{region 'Documentation'}
(*!
<summary>No asynchronous test resource remains to stop.</summary>
*)
{endregion}
METHOD PROTECTED ProcessAbort
VAR_INPUT
    Enable : BOOL; //! Phase permission supplied by the owning Test Case; FALSE does not authorize progression, while observation may continue.
END_VAR
IF Enable THEN
    CompleteAbort();
END_IF;
END_METHOD

{region 'Documentation'}
(*!
<summary>Evaluates each scripted call before the test advances; failures remain latched across both runs.</summary>
*)
{endregion}
METHOD PROTECTED ProcessAssertions
VAR_INPUT
    Enable : BOOL; //! Phase permission supplied by the owning Test Case; FALSE does not authorize progression, while observation may continue.
END_VAR
FStatePath(Enable := Enable,
    State := State,
    IN := FStatePathMatches);
FTaskMapping(Enable := Enable,
    State := State,
    IN := FTaskMappingMatches);
FOwnerResult(Enable := Enable,
    State := State,
    IN := FOwnerResultMatches);
FStatusCounters(Enable := Enable,
    State := State,
    IN := FStatusCountersMatches);
FCallOrder(Enable := Enable,
    State := State,
    IN := FCallOrderMatches);
FReadiness(Enable := Enable,
    State := State,
    IN := FReadinessMatches);
FFinalEvents(Enable := Enable,
    State := State,
    IN := FFinalEventsMatches);
FAggregationPayload(Enable := Enable,
    State := State,
    IN := FAggregationPayloadMatches);
FCaptureIntegrity(Enable := Enable,
    State := State,
    IN := FCaptureIntegrityMatches);
IF Enable THEN
    FStepChecked := TRUE;
END_IF;
END_METHOD

{region 'Documentation'}
(*!
<summary>No resource Preparation is required for this controlled owner scenario.</summary>
*)
{endregion}
METHOD PROTECTED ProcessPreparations
VAR_INPUT
    // SA0033: Required override; the scenario has no Preparation phase.
    {attribute 'analysis' := '-33'}
    Enable : BOOL; //! Phase permission supplied by the owning Test Case; FALSE does not authorize progression, while observation may continue.
END_VAR
END_METHOD

{region 'Documentation'}
(*!
<summary>Restarts the test script and clears checking Assertions; subject setup belongs to the next test attempt.</summary>
*)
{endregion}
METHOD PROTECTED ProcessReset
FStep := Setup;
FRun := 1;
FStepChecked := FALSE;
FStatePathMatches := TRUE;
FTaskMappingMatches := TRUE;
FOwnerResultMatches := TRUE;
FStatusCountersMatches := TRUE;
FCallOrderMatches := TRUE;
FReadinessMatches := TRUE;
FFinalEventsMatches := TRUE;
FAggregationPayloadMatches := TRUE;
FCaptureIntegrityMatches := TRUE;
FStatePath.Reset();
FTaskMapping.Reset();
FOwnerResult.Reset();
FStatusCounters.Reset();
FCallOrder.Reset();
FReadiness.Reset();
FFinalEvents.Reset();
FAggregationPayload.Reset();
FCaptureIntegrity.Reset();
CompleteReset();
END_METHOD

{region 'Documentation'}
(*!
<summary>Advances the explicit test script with at most one subject FB call per active PLC cycle.</summary>
*)
{endregion}
METHOD PROTECTED ProcessTests
VAR_INPUT
    Enable : BOOL; //! Phase permission supplied by the owning Test Case; FALSE does not authorize progression, while observation may continue.
END_VAR
IF NOT Enable THEN
    RETURN;
END_IF;
IF FStepChecked THEN
    IF FStep = StartWithoutReset THEN
        IF FRun = RunCount THEN
            CompleteTests();
            RETURN;
        END_IF;
        FRun := FRun + 1;
        FStep := Setup;
    ELSE
        FStep := FStep + 1;
    END_IF;
    FStepChecked := FALSE;
    NextTestState();
END_IF;
RunStep();
END_METHOD

{region 'Documentation'}
(*!
<summary>Arranges one root cycle, executes it once and compares state, counters and call ordering.</summary>
*)
{endregion}
METHOD PRIVATE RunStep
VAR
    Config : ST_RunConfig;
    FirstView : ST_OrchestrationObservation;
    SecondView : ST_OrchestrationObservation;
    ExpectedState : E_State;
    ExpectedTask : E_OrchestratorTask;
    ExpectedResult : E_Result := E_Result.NotEvaluated;
    ExpectedReady : BOOL;
    ExpectedIdleCount : UINT;
    ExpectedRunningCount : UINT;
    ExpectedCompletedCount : UINT;
    ExpectedPassedCount : UINT;
    ExpectedFailedCount : UINT;
    ExpectedExecutionStatus : E_ExecutionStatus;
    FirstChild : I_Orchestratable;
    LastChild : I_Orchestratable;
    FirstStateBeforeCall : E_State;
    LastStateBeforeCall : E_State;
    Snapshot : ST_RunControlStatus;
    ExpectedCalls : UINT;
END_VAR
CASE FStep OF
    Setup:
        FRunChildResult := E_Result.Passed;
        IF FRun = 1 THEN
            FRunChildResult := FirstChildResult;
            IF NOT FCapture.Initialize(Buffer := FEvents,
                FifoControl := FCaptureFifo,
                Status := FCaptureStatus) THEN
                Error(Message := 'Root lifecycle capture could not be initialized.');
                RETURN;
            END_IF;
            Config.CompletionDelay := T#0ms;
            FHelper.BeginScenario();
            FSubject.Bind(Publisher := FCapture,
                Helper := FHelper,
                Config := Config);
            IF NOT FSubject.Initialize(Name := 'LifecycleSubject',
                EventBuffer := FCapture) THEN
                Error(Message := 'Root lifecycle subject could not be initialized.');
                RETURN;
            END_IF;
        ELSE
            FHelper.SetObservation(Ready := FALSE);
            FSubject.RequestReset();
        END_IF;
        FirstView.State := E_State.Reset;
        FirstView.Ready := FALSE;
        SecondView := FirstView;
        ExpectedState := E_State.Reset;
        ExpectedTask := E_OrchestratorTask.Reset;
        ExpectedExecutionStatus := E_ExecutionStatus.Reset;

    ChildrenReady:
        ExpectedState := E_State.Reset;
        ExpectedTask := E_OrchestratorTask.Reset;
        ExpectedExecutionStatus := E_ExecutionStatus.Reset;
        ExpectedIdleCount := ExpectedChildCount;

    ResetFinished:
        FHelper.SetObservation(Ready := FALSE,
            ResetFinished := TRUE);
        ExpectedState := E_State.Idle;
        ExpectedTask := E_OrchestratorTask.Idle;
        ExpectedExecutionStatus := E_ExecutionStatus.Idle;
        ExpectedIdleCount := ExpectedChildCount;

    StartReady:
        FHelper.SetObservation(Ready := TRUE);
        ExpectedState := E_State.Idle;
        ExpectedTask := E_OrchestratorTask.Idle;
        ExpectedExecutionStatus := E_ExecutionStatus.Idle;
        ExpectedIdleCount := ExpectedChildCount;
        ExpectedReady := TRUE;

    StartRequested:
        FSubject.RequestStart();
        FirstView.State := E_State.Running;
        FirstView.Ready := FALSE;
        ExpectedState := E_State.Starting;
        ExpectedTask := E_OrchestratorTask.Execution;
        ExpectedExecutionStatus := E_ExecutionStatus.Starting;
        ExpectedIdleCount := 1;
        ExpectedRunningCount := 1;

    FirstChildCompleted:
        FHelper.SetObservation(Ready := FALSE);
        FirstView.State := E_State.Completed;
        FirstView.Result := FRunChildResult;
        FirstView.Ready := FALSE;
        FirstView.Complete := TRUE;
        SecondView.State := E_State.Running;
        SecondView.Ready := FALSE;
        ExpectedState := E_State.Running;
        ExpectedTask := E_OrchestratorTask.Execution;
        ExpectedExecutionStatus := E_ExecutionStatus.Running;
        ExpectedRunningCount := 1;
        ExpectedCompletedCount := 1;
        ExpectedFailedCount := BOOL_TO_UINT(FRunChildResult = E_Result.Failed);
        ExpectedPassedCount := 1 - ExpectedFailedCount;

    AllChildrenCompleted, WaitForHelper, OwnerCompleting, OwnerCompleted, HoldCompleted, StartWithoutReset:
        FHelper.SetObservation(Ready := FALSE);
        FirstView.State := E_State.Completed;
        FirstView.Result := FRunChildResult;
        FirstView.Ready := FALSE;
        FirstView.Complete := TRUE;
        SecondView := FirstView;
        SecondView.Result := E_Result.Passed;
        ExpectedTask := E_OrchestratorTask.Execution;
        ExpectedCompletedCount := ExpectedChildCount;
        ExpectedFailedCount := BOOL_TO_UINT(FRunChildResult = E_Result.Failed);
        ExpectedPassedCount := ExpectedChildCount - ExpectedFailedCount;
        CASE FStep OF
            AllChildrenCompleted, WaitForHelper:
                ExpectedState := E_State.Running;
                ExpectedExecutionStatus := E_ExecutionStatus.Running;
            OwnerCompleting:
                FHelper.SetObservation(Ready := FALSE,
                    ExecutionFinished := TRUE);
                ExpectedState := E_State.Completing;
                ExpectedExecutionStatus := E_ExecutionStatus.Completing;
                ExpectedResult := FRunChildResult;
        ELSE
            IF FStep = StartWithoutReset THEN
                FSubject.RequestStart();
            END_IF;
            ExpectedState := E_State.Completed;
            ExpectedTask := E_OrchestratorTask.Idle;
            ExpectedExecutionStatus := E_ExecutionStatus.Completed;
            ExpectedResult := FRunChildResult;
        END_CASE;
ELSE
    Error(Message := 'Unexpected root lifecycle test step.');
    RETURN;
END_CASE;

FirstChild := FSubject.GetChild(Index := FSubject.ChildArrayLowerBound);
LastChild := FSubject.GetChild(Index := FSubject.ChildArrayLowerBound + UINT_TO_DINT(FSubject.ChildCount) - 1);
FirstStateBeforeCall := FirstChild.State;
LastStateBeforeCall := LastChild.State;
FSubject.SetChildObservations(FirstChild := FirstView,
    SecondChild := SecondView);
FSubject(ControlData := FControl);
Snapshot := FSubject.Status;
ExpectedCalls := INT_TO_UINT((FRun - 1) * StepsPerRun + FStep + 1);

FStatePathMatches := (FSubject.State = ExpectedState)
    AND (Snapshot.Execution.State = ExpectedState)
    AND (Snapshot.Execution.ExecutionStatus = ExpectedExecutionStatus)
    AND (FControl.Status.Execution.State = ExpectedState)
    AND (FControl.Name = 'LifecycleSubject');
FTaskMappingMatches := FHelper.CurrentTask = ExpectedTask;
FOwnerResultMatches := (FSubject.Result = ExpectedResult)
    AND (Snapshot.Execution.Result = ExpectedResult)
    AND (FControl.Status.Execution.Result = ExpectedResult)
    AND NOT FSubject.HasError;
FStatusCountersMatches := (Snapshot.SuiteCountTotal = ExpectedChildCount)
    AND (Snapshot.SuiteCountIdle = ExpectedIdleCount)
    AND (Snapshot.SuiteCountRunning = ExpectedRunningCount)
    AND (Snapshot.SuiteCountCompleted = ExpectedCompletedCount)
    AND (Snapshot.SuiteCountPassed = ExpectedPassedCount)
    AND (Snapshot.SuiteCountFailed = ExpectedFailedCount)
    AND (Snapshot.SuiteCountError = 0) AND (Snapshot.SuiteCountInactive = 0)
    AND (FControl.Status.SuiteCountIdle = ExpectedIdleCount)
    AND (FControl.Status.SuiteCountRunning = ExpectedRunningCount)
    AND (FControl.Status.SuiteCountCompleted = ExpectedCompletedCount)
    AND (FControl.Status.SuiteCountPassed = ExpectedPassedCount)
    AND (FControl.Status.SuiteCountFailed = ExpectedFailedCount);
FCallOrderMatches := (FHelper.InitializeCount = 1) AND (FSubject.ConfigureCount = 1)
    AND (FHelper.ExecuteCount = ExpectedCalls)
    AND (FSubject.ChildCallCount = ExpectedCalls)
    AND FSubject.ChildBodyCallsMatch
    AND (FHelper.FirstChildStateAtExecute = FirstStateBeforeCall)
    AND (FHelper.LastChildStateAtExecute = LastStateBeforeCall)
    AND (FirstChild.State = FirstView.State) AND (LastChild.State = SecondView.State);
FReadinessMatches := (FSubject.IsReady = ExpectedReady)
    AND (Snapshot.Execution.Ready = ExpectedReady)
    AND (FSubject.IsComplete = (ExpectedState = E_State.Completed));
FCaptureIntegrityMatches := (FCaptureStatus.LostEventCount = 0)
    AND (FCaptureFifo.ElementCount = FCaptureStatus.SequenceId);
IF FStep = Setup THEN
    FOwnerResultMatches := FOwnerResultMatches AND (Snapshot.Runtime = T#0ms);
END_IF;
IF FStep = OwnerCompleting THEN
    FRunRuntime[FRun] := Snapshot.Runtime;
END_IF;
CheckFinalEvents();
END_METHOD

END_FUNCTION_BLOCK

// ---- SelfTests/TestCases/TestSuite_RunControlLifecycle/Test_RunControlRequests.TcPOU
{region 'Documentation'}
(*!
<summary>Checks direct root requests, one-call consumption and Reset/Abort/Start priority.</summary>
<description>
The controlled helper only supplies readiness and completion. The script covers a Start
received while not ready, repeated Start method calls before one FB call, Start while active,
Abort together with Start, and Reset together with both lower-priority requests.
A repeated Reset while already resetting still has one trigger but no repeated transition.
Following request-free calls verify that consumed requests cannot replay.
Checks before the subject call prove that the methods do not advance its lifecycle or publish.
The active Reset warning is expected and isolated; this scenario never finalizes a run.
External command bits and their two-sample qualification are deliberately not exercised.
</description>
*)
{endregion}
FUNCTION_BLOCK Test_RunControlRequests EXTENDS TestCaseBase
VAR
    FSubject : RunControlLifecycleProbe;
    FHelper : SuiteOrchestratorDouble;
    FControl : ST_RunControl;
    FCapture : EventBuffer;
    FEvents : ARRAY[1..CaptureLength] OF ST_Event;
    FCaptureFifo : ST_FifoStatus;
    FCaptureStatus : ST_EventBufferStatus;
    FStep : INT;
    FStepChecked : BOOL;
    FLifecycle : AssertTrue;
    FLifecycleMatches : BOOL := TRUE;
    FDeferredRequests : AssertTrue;
    FDeferredRequestsMatches : BOOL := TRUE;
    FTriggerEvidence : AssertTrue;
    FTriggerEvidenceMatches : BOOL := TRUE;
    FEventBoundary : AssertTrue;
    FEventBoundaryMatches : BOOL := TRUE;
    FProjection : AssertTrue;
    FProjectionMatches : BOOL := TRUE;
    FDispatch : AssertTrue;
    FDispatchMatches : BOOL := TRUE;
END_VAR
VAR CONSTANT
    CaptureLength : UINT := 64;
    Setup : INT := 0;
    InitialIdle : INT := 1;
    StartNotReady : INT := 2;
    ReadyWithoutRequest : INT := 3;
    RepeatedStart : INT := 4;
    StartWhileActive : INT := 5;
    AbortOverStart : INT := 6;
    ResetOverAll : INT := 7;
    RepeatReset : INT := 8;
    ResetFinished : INT := 9;
    NoReplayAfterReset : INT := 10;
    AbortInIdle : INT := 11;
    NoReplayAfterAbort : INT := 12;
    StepCount : INT := 13;
END_VAR

SUPER^();

{region 'Documentation'}
(*!
<summary>Contributes only the checking Assertions, not the intentionally controlled subject results.</summary>
*)
{endregion}
METHOD PROTECTED AggregateResults
VAR_INPUT
    Aggregator : I_ResultAggregator; //! Borrowed result sink owned by the outer Test Case; add this test's checking Assertions without resetting or retaining the sink.
END_VAR
Aggregator.AddProvider(Provider := FLifecycle);
Aggregator.AddProvider(Provider := FDeferredRequests);
Aggregator.AddProvider(Provider := FTriggerEvidence);
Aggregator.AddProvider(Provider := FEventBoundary);
Aggregator.AddProvider(Provider := FProjection);
Aggregator.AddProvider(Provider := FDispatch);
END_METHOD

{region 'Documentation'}
(*!
<summary>Initializes the checking Assertions; the scenario explicitly initializes its isolated subject.</summary>
*)
{endregion}
METHOD PROTECTED Configure
FPreparationStateCount := 0;
FTestStateCount := StepCount;
FLifecycle.Initialize(Parent := THIS^,
    AssertionName := 'Lifecycle');
FDeferredRequests.Initialize(Parent := THIS^,
    AssertionName := 'DeferredRequests');
FTriggerEvidence.Initialize(Parent := THIS^,
    AssertionName := 'TriggerEvidence');
FEventBoundary.Initialize(Parent := THIS^,
    AssertionName := 'EventBoundary');
FProjection.Initialize(Parent := THIS^,
    AssertionName := 'Projection');
FDispatch.Initialize(Parent := THIS^,
    AssertionName := 'Dispatch');
END_METHOD

{region 'Documentation'}
(*!
<summary>No asynchronous test resource remains to stop.</summary>
*)
{endregion}
METHOD PROTECTED ProcessAbort
VAR_INPUT
    Enable : BOOL; //! Phase permission supplied by the owning Test Case; FALSE does not authorize progression, while observation may continue.
END_VAR
IF Enable THEN
    CompleteAbort();
END_IF;
END_METHOD

{region 'Documentation'}
(*!
<summary>Checks each request step before advancing; no expected subject result is counted as a test Assertion.</summary>
*)
{endregion}
METHOD PROTECTED ProcessAssertions
VAR_INPUT
    Enable : BOOL; //! Phase permission supplied by the owning Test Case; FALSE does not authorize progression, while observation may continue.
END_VAR
FLifecycle(Enable := Enable,
    State := State,
    IN := FLifecycleMatches);
FDeferredRequests(Enable := Enable,
    State := State,
    IN := FDeferredRequestsMatches);
FTriggerEvidence(Enable := Enable,
    State := State,
    IN := FTriggerEvidenceMatches);
FEventBoundary(Enable := Enable,
    State := State,
    IN := FEventBoundaryMatches);
FProjection(Enable := Enable,
    State := State,
    IN := FProjectionMatches);
FDispatch(Enable := Enable,
    State := State,
    IN := FDispatchMatches);
IF Enable THEN
    FStepChecked := TRUE;
END_IF;
END_METHOD

{region 'Documentation'}
(*!
<summary>No resource Preparation is required for this controlled owner scenario.</summary>
*)
{endregion}
METHOD PROTECTED ProcessPreparations
VAR_INPUT
    // SA0033: Required override; the scenario has no Preparation phase.
    {attribute 'analysis' := '-33'}
    Enable : BOOL; //! Phase permission supplied by the owning Test Case; FALSE does not authorize progression, while observation may continue.
END_VAR
END_METHOD

{region 'Documentation'}
(*!
<summary>Restarts the test script and clears checking Assertions; subject setup belongs to the next test attempt.</summary>
*)
{endregion}
METHOD PROTECTED ProcessReset
FStep := Setup;
FStepChecked := FALSE;
FLifecycleMatches := TRUE;
FDeferredRequestsMatches := TRUE;
FTriggerEvidenceMatches := TRUE;
FEventBoundaryMatches := TRUE;
FProjectionMatches := TRUE;
FDispatchMatches := TRUE;
FLifecycle.Reset();
FDeferredRequests.Reset();
FTriggerEvidence.Reset();
FEventBoundary.Reset();
FProjection.Reset();
FDispatch.Reset();
CompleteReset();
END_METHOD

{region 'Documentation'}
(*!
<summary>Advances the explicit test script with at most one subject FB call per active PLC cycle.</summary>
*)
{endregion}
METHOD PROTECTED ProcessTests
VAR_INPUT
    Enable : BOOL; //! Phase permission supplied by the owning Test Case; FALSE does not authorize progression, while observation may continue.
END_VAR
IF NOT Enable THEN
    RETURN;
END_IF;
IF FStepChecked THEN
    IF FStep = NoReplayAfterAbort THEN
        CompleteTests();
        RETURN;
    END_IF;
    FStep := FStep + 1;
    FStepChecked := FALSE;
    NextTestState();
END_IF;
RunStep();
END_METHOD

{region 'Documentation'}
(*!
<summary>Applies direct requests before one subject call; counts semantic event types, never diagnostic wording.</summary>
*)
{endregion}
METHOD PRIVATE RunStep
VAR
    Config : ST_RunConfig;
    ChildView : ST_OrchestrationObservation;
    ExpectedState : E_State := E_State.Idle;
    ExpectedTask : E_OrchestratorTask := E_OrchestratorTask.Idle;
    ExpectedResult : E_Result := E_Result.NotEvaluated;
    ExpectedReady : BOOL;
    ExpectedTriggers : UINT;
    ExpectedWarnings : UINT;
    TriggerCount : UINT;
    WarningCount : UINT;
    Index : UINT;
    StateBeforeRequest : E_State;
    ResultBeforeRequest : E_Result;
    SequenceBeforeRequest : UDINT;
    SequenceBeforeCall : UDINT;
END_VAR
IF FStep = Setup THEN
    IF NOT FCapture.Initialize(Buffer := FEvents,
        FifoControl := FCaptureFifo,
        Status := FCaptureStatus) THEN
        Error(Message := 'Root request capture could not be initialized.');
        RETURN;
    END_IF;
    FHelper.BeginScenario();
    FSubject.Bind(Publisher := FCapture,
        Helper := FHelper,
        Config := Config);
    IF NOT FSubject.Initialize(Name := 'RequestSubject',
        EventBuffer := FCapture) THEN
        Error(Message := 'Root request subject could not be initialized.');
        RETURN;
    END_IF;
END_IF;

StateBeforeRequest := FSubject.State;
ResultBeforeRequest := FSubject.Result;
SequenceBeforeRequest := FCaptureStatus.SequenceId;
FHelper.SetObservation(Ready := FALSE);
CASE FStep OF
    Setup:
        ExpectedState := E_State.Reset;
        ExpectedTask := E_OrchestratorTask.Reset;
        ExpectedTriggers := 1;
    InitialIdle:
        FHelper.SetObservation(Ready := TRUE,
            ResetFinished := TRUE);
        ExpectedReady := TRUE;
        ExpectedTriggers := 1;
    StartNotReady:
        FSubject.RequestStart();
        ExpectedTriggers := 2;
    ReadyWithoutRequest:
        FHelper.SetObservation(Ready := TRUE);
        ExpectedReady := TRUE;
        ExpectedTriggers := 2;
    RepeatedStart:
        FHelper.SetObservation(Ready := TRUE);
        FSubject.RequestStart();
        FSubject.RequestStart();
        ChildView.State := E_State.Running;
        ChildView.Ready := FALSE;
        ExpectedState := E_State.Starting;
        ExpectedTask := E_OrchestratorTask.Execution;
        ExpectedTriggers := 3;
    StartWhileActive:
        FSubject.RequestStart();
        ChildView.State := E_State.Running;
        ChildView.Ready := FALSE;
        ExpectedState := E_State.Running;
        ExpectedTask := E_OrchestratorTask.Execution;
        ExpectedTriggers := 4;
    AbortOverStart:
        FSubject.RequestStart();
        FSubject.RequestAbort();
        ChildView.State := E_State.Running;
        ChildView.Ready := FALSE;
        ExpectedState := E_State.Aborting;
        ExpectedTask := E_OrchestratorTask.Abort;
        ExpectedResult := E_Result.Abort;
        ExpectedTriggers := 6;
    ResetOverAll:
        FSubject.RequestStart();
        FSubject.RequestAbort();
        FSubject.RequestReset();
        ChildView.State := E_State.Reset;
        ChildView.Ready := FALSE;
        ExpectedState := E_State.Reset;
        ExpectedTask := E_OrchestratorTask.Reset;
        ExpectedTriggers := 9;
    RepeatReset:
        FSubject.RequestReset();
        ExpectedState := E_State.Reset;
        ExpectedTask := E_OrchestratorTask.Reset;
        ExpectedTriggers := 10;
    ResetFinished:
        FHelper.SetObservation(Ready := TRUE,
            ResetFinished := TRUE);
        ExpectedReady := TRUE;
        ExpectedTriggers := 10;
    NoReplayAfterReset:
        FHelper.SetObservation(Ready := TRUE);
        ExpectedReady := TRUE;
        ExpectedTriggers := 10;
    AbortInIdle, NoReplayAfterAbort:
        IF FStep = AbortInIdle THEN
            FSubject.RequestAbort();
        END_IF;
        FHelper.SetObservation(Ready := TRUE);
        ExpectedReady := TRUE;
        ExpectedTriggers := 11;
ELSE
    Error(Message := 'Unexpected root request test step.');
    RETURN;
END_CASE;
FDeferredRequestsMatches := (FSubject.State = StateBeforeRequest)
    AND (FSubject.Result = ResultBeforeRequest)
    AND (FCaptureStatus.SequenceId = SequenceBeforeRequest);
SequenceBeforeCall := FCaptureStatus.SequenceId;
FSubject.SetChildObservation(Observation := ChildView);
FSubject(ControlData := FControl);
FLifecycleMatches := (FSubject.State = ExpectedState)
    AND (FSubject.Result = ExpectedResult)
    AND (FSubject.IsReady = ExpectedReady)
    AND (FHelper.CurrentTask = ExpectedTask)
    AND NOT FSubject.HasError;
FProjectionMatches := (FControl.Name = 'RequestSubject')
    AND (FControl.Status.Execution.State = ExpectedState)
    AND (FControl.Status.Execution.Result = ExpectedResult)
    AND (FControl.Status.Execution.Ready = ExpectedReady);
FDispatchMatches := (FHelper.ExecuteCount = INT_TO_UINT(FStep + 1))
    AND (FSubject.ChildCallCount = INT_TO_UINT(FStep + 1))
    AND FSubject.ChildBodyCallsMatch
    AND (FHelper.InitializeCount = 1) AND (FSubject.ConfigureCount = 1);

FEventBoundaryMatches := TRUE;
FOR Index := 1 TO FCaptureFifo.ElementCount DO
    FEventBoundaryMatches := FEventBoundaryMatches
        AND (FEvents[Index].OwnerScope = E_OwnerScope.RunControl)
        AND (FEvents[Index].Name = 'RequestSubject')
        AND (FEvents[Index].EventType <> E_EventType.Result)
        AND (FEvents[Index].EventType <> E_EventType.Aggregation)
        AND (FEvents[Index].Severity <> E_EventSeverity.Error);
    IF FEvents[Index].EventType = E_EventType.Trigger THEN
        TriggerCount := TriggerCount + 1;
    END_IF;
    IF FEvents[Index].Severity = E_EventSeverity.Warning THEN
        WarningCount := WarningCount + 1;
    END_IF;
END_FOR;
ExpectedWarnings := BOOL_TO_UINT(FStep >= ResetOverAll);
FEventBoundaryMatches := FEventBoundaryMatches
    AND (WarningCount = ExpectedWarnings)
    AND (FCaptureStatus.LostEventCount = 0);
FTriggerEvidenceMatches := TriggerCount = ExpectedTriggers;
IF FStep = RepeatReset THEN
    FTriggerEvidenceMatches := FTriggerEvidenceMatches
        AND (FCaptureStatus.SequenceId = SequenceBeforeCall + 1);
END_IF;
END_METHOD

END_FUNCTION_BLOCK

// ---- SelfTests/TestCases/TestSuite_RunControlLifecycle/Test_RunControlRealComposition.TcPOU
{region 'Documentation'}
(*!
<summary>Runs the real root-to-Test-Case hierarchy twice with lifecycle Reset between executions.</summary>
<description>

Real boundaries

The local root owns a real Suite with two minimal real Test Cases. Both owner levels use
the production Orchestrator. The test supplies root Reset/Start requests only; scheduling
and every reservation/free operation belong to the real hierarchy.

Repeat and isolation

Initialize runs once. Two executions must finish Passed with lifecycle Reset between them.
Every producer uses one private Event Buffer retained across both executions. The outer
selftest runner remains unchanged. Child finalizations must precede their owner finalization,
and root completion must leave no reservations. Scheduling-mode matrices are not repeated.
</description>
*)
{endregion}
FUNCTION_BLOCK Test_RunControlRealComposition EXTENDS TestCaseBase
VAR
    FSubject : RunControlIntegrationSubject;
    FControl : ST_RunControl;
    FCapture : EventBuffer;
    FEvents : ARRAY[1..CaptureLength] OF ST_Event;
    FCaptureFifo : ST_FifoStatus;
    FCaptureStatus : ST_EventBufferStatus;
    FStep : INT;
    FCompletedRuns : UINT;
    FFinalChecksEvaluated : BOOL;
    FReadiness : AssertTrue;
    FReadinessMatches : BOOL := TRUE;
    FCompletion : AssertTrue;
    FCompletionMatches : BOOL := TRUE;
    FRepeat : AssertTrue;
    FRepeatMatches : BOOL := TRUE;
    FReservations : AssertTrue;
    FReservationsMatches : BOOL := TRUE;
    FChildCalls : AssertTrue;
    FChildCallsMatches : BOOL := TRUE;
    FEventStream : AssertTrue;
    FEventStreamMatches : BOOL := TRUE;
END_VAR
VAR CONSTANT
    CaptureLength : UINT := 512;
    ExpectedChildCount : UINT := 1;
    RequiredRuns : UINT := 2;
    Setup : INT := 0;
    ResetRequested : INT := 1;
    WaitForReadiness : INT := 2;
    StartRequested : INT := 3;
    WaitForCompletion : INT := 4;
    Finish : INT := 5;
END_VAR

SUPER^();

{region 'Documentation'}
(*!
<summary>Contributes only the checking Assertions, not the intentionally controlled subject results.</summary>
*)
{endregion}
METHOD PROTECTED AggregateResults
VAR_INPUT
    Aggregator : I_ResultAggregator; //! Borrowed result sink owned by the outer Test Case; add this test's checking Assertions without resetting or retaining the sink.
END_VAR
Aggregator.AddProvider(Provider := FReadiness);
Aggregator.AddProvider(Provider := FCompletion);
Aggregator.AddProvider(Provider := FRepeat);
Aggregator.AddProvider(Provider := FReservations);
Aggregator.AddProvider(Provider := FChildCalls);
Aggregator.AddProvider(Provider := FEventStream);
END_METHOD

{region 'Documentation'}
(*!
<summary>Checks exact finalization counts and latest child-before-owner event order across both executions.</summary>
*)
{endregion}
METHOD PRIVATE CheckEventStream
VAR
    Index : UINT;
    Suite : I_TestSuite;
    RootResults : UINT;
    RootAggregations : UINT;
    RootCompletions : UINT;
    RootResultSequence : UDINT;
    RootAggregationSequence : UDINT;
    RootCompletionSequence : UDINT;
    SuiteResults : UINT;
    SuiteAggregations : UINT;
    SuiteCompletions : UINT;
    FirstResults : UINT;
    SecondResults : UINT;
    FirstCompletions : UINT;
    SecondCompletions : UINT;
    SuiteResultSequence : UDINT;
    SuiteAggregationSequence : UDINT;
    SuiteCompletionSequence : UDINT;
    FirstCompletionSequence : UDINT;
    SecondCompletionSequence : UDINT;
    FirstChild : I_TestCase;
    SecondChild : I_TestCase;
END_VAR
Suite := FSubject.GetTestSuite(Index := FSubject.ChildArrayLowerBound);
FirstChild := FSubject.GetTestCase(Index := FSubject.TestCaseLowerBound);
SecondChild := FSubject.GetTestCase(Index := FSubject.TestCaseLowerBound + 1);
FOR Index := 1 TO CaptureLength DO
    IF FEvents[Index].SequenceId = 0 THEN
        CONTINUE;
    END_IF;
    FEventStreamMatches := FEventStreamMatches
        AND (FEvents[Index].Severity <> E_EventSeverity.Error);
    IF FEvents[Index].Name = FSubject.Name THEN
        CASE FEvents[Index].EventType OF
            E_EventType.Result:
                RootResults := RootResults + 1;
                RootResultSequence := FEvents[Index].SequenceId;
                FEventStreamMatches := FEventStreamMatches AND (FEvents[Index].Result = E_Result.Passed)
                    AND (FEvents[Index].OwnerScope = E_OwnerScope.RunControl);
            E_EventType.Aggregation:
                RootAggregations := RootAggregations + 1;
                RootAggregationSequence := FEvents[Index].SequenceId;
            E_EventType.StateTransition:
                IF FEvents[Index].State = E_State.Completed THEN
                    RootCompletions := RootCompletions + 1;
                    RootCompletionSequence := FEvents[Index].SequenceId;
                END_IF;
        END_CASE;
    ELSIF FEvents[Index].Name = Suite.Name THEN
        CASE FEvents[Index].EventType OF
            E_EventType.Result:
                SuiteResults := SuiteResults + 1;
                SuiteResultSequence := FEvents[Index].SequenceId;
                FEventStreamMatches := FEventStreamMatches AND (FEvents[Index].Result = E_Result.Passed);
            E_EventType.Aggregation:
                SuiteAggregations := SuiteAggregations + 1;
                SuiteAggregationSequence := FEvents[Index].SequenceId;
            E_EventType.StateTransition:
                IF FEvents[Index].State = E_State.Completed THEN
                    SuiteCompletions := SuiteCompletions + 1;
                    SuiteCompletionSequence := FEvents[Index].SequenceId;
                END_IF;
        END_CASE;
    ELSIF FEvents[Index].Name = FirstChild.Name THEN
        IF FEvents[Index].EventType = E_EventType.Result THEN
            FirstResults := FirstResults + 1;
        ELSIF (FEvents[Index].EventType = E_EventType.StateTransition)
            AND (FEvents[Index].State = E_State.Completed) THEN
            FirstCompletions := FirstCompletions + 1;
            FirstCompletionSequence := FEvents[Index].SequenceId;
        END_IF;
    ELSIF FEvents[Index].Name = SecondChild.Name THEN
        IF FEvents[Index].EventType = E_EventType.Result THEN
            SecondResults := SecondResults + 1;
        ELSIF (FEvents[Index].EventType = E_EventType.StateTransition)
            AND (FEvents[Index].State = E_State.Completed) THEN
            SecondCompletions := SecondCompletions + 1;
            SecondCompletionSequence := FEvents[Index].SequenceId;
        END_IF;
    END_IF;
END_FOR;
FEventStreamMatches := FEventStreamMatches
    AND (SuiteResults = FCompletedRuns) AND (SuiteAggregations = FCompletedRuns)
    AND (SuiteCompletions = FCompletedRuns)
    AND (FirstResults = FCompletedRuns) AND (SecondResults = FCompletedRuns)
    AND (FirstCompletions = FCompletedRuns) AND (SecondCompletions = FCompletedRuns)
    AND (FirstCompletionSequence < SuiteResultSequence)
    AND (SecondCompletionSequence < SuiteResultSequence)
    AND (SuiteResultSequence < SuiteAggregationSequence)
    AND (SuiteAggregationSequence < SuiteCompletionSequence)
    AND (RootResults = FCompletedRuns) AND (RootAggregations = FCompletedRuns)
    AND (RootCompletions = FCompletedRuns)
    AND (SuiteCompletionSequence < RootResultSequence)
    AND (RootResultSequence < RootAggregationSequence)
    AND (RootAggregationSequence < RootCompletionSequence);
END_METHOD

{region 'Documentation'}
(*!
<summary>Observes cleanup performed by the real hierarchy; the test does not release any reservation.</summary>
*)
{endregion}
METHOD PRIVATE CheckReservations
VAR
    Suite : I_TestSuite;
    FirstChild : I_TestCase;
    SecondChild : I_TestCase;
END_VAR
Suite := FSubject.GetTestSuite(Index := FSubject.ChildArrayLowerBound);
FirstChild := FSubject.GetTestCase(Index := FSubject.TestCaseLowerBound);
SecondChild := FSubject.GetTestCase(Index := FSubject.TestCaseLowerBound + 1);
FReservationsMatches := FReservationsMatches
    AND (Suite.ReservedEntryCount = 0)
    AND (FirstChild.ReservedEntryCount = 0) AND (SecondChild.ReservedEntryCount = 0)
    AND (FCapture.ReservedEntryCount = 0);
END_METHOD

{region 'Documentation'}
(*!
<summary>Initializes the checking Assertions; the scenario explicitly initializes its isolated subject.</summary>
*)
{endregion}
METHOD PROTECTED Configure
FPreparationStateCount := 0;
FTestStateCount := 1;
FReadiness.Initialize(Parent := THIS^,
    AssertionName := 'Readiness');
FCompletion.Initialize(Parent := THIS^,
    AssertionName := 'Completion');
FRepeat.Initialize(Parent := THIS^,
    AssertionName := 'Repeat');
FReservations.Initialize(Parent := THIS^,
    AssertionName := 'Reservations');
FChildCalls.Initialize(Parent := THIS^,
    AssertionName := 'ChildCalls');
FEventStream.Initialize(Parent := THIS^,
    AssertionName := 'EventStream');
END_METHOD

{region 'Documentation'}
(*!
<summary>No asynchronous test resource remains to stop.</summary>
*)
{endregion}
METHOD PROTECTED ProcessAbort
VAR_INPUT
    Enable : BOOL; //! Phase permission supplied by the owning Test Case; FALSE does not authorize progression, while observation may continue.
END_VAR
IF Enable THEN
    CompleteAbort();
END_IF;
END_METHOD

{region 'Documentation'}
(*!
<summary>Keeps every observation across both runs; final checks must evaluate before ending the outer Test Case.</summary>
*)
{endregion}
METHOD PROTECTED ProcessAssertions
VAR_INPUT
    Enable : BOOL; //! Phase permission supplied by the owning Test Case; FALSE does not authorize progression, while observation may continue.
END_VAR
FReadiness(Enable := Enable,
    State := State,
    IN := FReadinessMatches);
FCompletion(Enable := Enable,
    State := State,
    IN := FCompletionMatches);
FRepeat(Enable := Enable,
    State := State,
    IN := FRepeatMatches);
FReservations(Enable := Enable,
    State := State,
    IN := FReservationsMatches);
FChildCalls(Enable := Enable,
    State := State,
    IN := FChildCallsMatches);
FEventStream(Enable := Enable,
    State := State,
    IN := FEventStreamMatches);
IF Enable AND (FStep = Finish) THEN
    FFinalChecksEvaluated := TRUE;
END_IF;
END_METHOD

{region 'Documentation'}
(*!
<summary>No resource Preparation is required for this controlled owner scenario.</summary>
*)
{endregion}
METHOD PROTECTED ProcessPreparations
VAR_INPUT
    // SA0033: Required override; the scenario has no Preparation phase.
    {attribute 'analysis' := '-33'}
    Enable : BOOL; //! Phase permission supplied by the owning Test Case; FALSE does not authorize progression, while observation may continue.
END_VAR
END_METHOD

{region 'Documentation'}
(*!
<summary>Restarts the test script and clears checking Assertions; subject setup belongs to the next test attempt.</summary>
*)
{endregion}
METHOD PROTECTED ProcessReset
FStep := Setup;
FCompletedRuns := 0;
FFinalChecksEvaluated := FALSE;
FReadinessMatches := TRUE;
FCompletionMatches := TRUE;
FRepeatMatches := TRUE;
FReservationsMatches := TRUE;
FChildCallsMatches := TRUE;
FEventStreamMatches := TRUE;
FReadiness.Reset();
FCompletion.Reset();
FRepeat.Reset();
FReservations.Reset();
FChildCalls.Reset();
FEventStream.Reset();
CompleteReset();
END_METHOD

{region 'Documentation'}
(*!
<summary>Advances the explicit test script with at most one subject FB call per active PLC cycle.</summary>
*)
{endregion}
METHOD PROTECTED ProcessTests
VAR_INPUT
    Enable : BOOL; //! Phase permission supplied by the owning Test Case; FALSE does not authorize progression, while observation may continue.
END_VAR
IF NOT Enable THEN
    RETURN;
END_IF;
IF (FStep = Finish) AND FFinalChecksEvaluated THEN
    CompleteTests();
    RETURN;
END_IF;
RunStep();
END_METHOD

{region 'Documentation'}
(*!
<summary>Issues root requests once; all lower-level requests and reservation handling remain production behavior.</summary>
*)
{endregion}
METHOD PRIVATE RunStep
VAR
    Snapshot : ST_RunControlStatus;
    Suite : I_TestSuite;
    FirstChild : I_TestCase;
    SecondChild : I_TestCase;
END_VAR
CASE FStep OF
    Setup:
        IF NOT FCapture.Initialize(Buffer := FEvents,
            FifoControl := FCaptureFifo,
            Status := FCaptureStatus) THEN
            Error(Message := 'Real root composition capture initialization failed.');
            RETURN;
        END_IF;
        FSubject.BindPublisher(Publisher := FCapture);
        IF NOT FSubject.Initialize(Name := 'RealRoot',
            EventBuffer := FCapture) THEN
            Error(Message := 'Real root composition initialization failed.');
            RETURN;
        END_IF;
        FStep := WaitForReadiness;

    ResetRequested:
        FSubject.RequestReset();
        FStep := WaitForReadiness;

    StartRequested:
        FSubject.RequestStart();
        FStep := WaitForCompletion;

    WaitForReadiness, WaitForCompletion, Finish:
        // The outer Test Case timeout bounds a stalled real hierarchy.
ELSE
    Error(Message := 'Unexpected real root composition test step.');
    RETURN;
END_CASE;

FSubject(ControlData := FControl);
FChildCallsMatches := FChildCallsMatches AND FSubject.ChildCallsMatch;
FRepeatMatches := FRepeatMatches AND FSubject.ConfigurationUnchanged
    AND (FSubject.ChildCount = ExpectedChildCount);
FEventStreamMatches := FEventStreamMatches AND (FCaptureStatus.LostEventCount = 0);
Snapshot := FSubject.Status;

CASE FStep OF
    WaitForReadiness:
        IF FSubject.HasError THEN
            Error(Message := 'Real root composition failed during Reset.');
            RETURN;
        END_IF;
        IF FSubject.IsReady THEN
            FReadinessMatches := FReadinessMatches AND FSubject.IsIdle
                AND (FSubject.Result = E_Result.NotEvaluated)
                AND (Snapshot.SuiteCountIdle = ExpectedChildCount)
                AND (Snapshot.SuiteCountCompleted = 0);
            CheckReservations();
            FStep := StartRequested;
        END_IF;

    WaitForCompletion:
        IF FSubject.IsComplete THEN
            Suite := FSubject.GetTestSuite(Index := FSubject.ChildArrayLowerBound);
            FirstChild := FSubject.GetTestCase(Index := FSubject.TestCaseLowerBound);
            SecondChild := FSubject.GetTestCase(Index := FSubject.TestCaseLowerBound + 1);
            FCompletionMatches := FCompletionMatches
                AND (FSubject.Result = E_Result.Passed)
                AND (FControl.Status.Execution.Result = E_Result.Passed)
                AND (Snapshot.SuiteCountCompleted = ExpectedChildCount)
                AND (Snapshot.SuiteCountPassed = ExpectedChildCount)
                AND (Snapshot.SuiteCountFailed = 0) AND (Snapshot.SuiteCountError = 0)
                AND Suite.IsComplete AND (Suite.Result = E_Result.Passed)
                AND FirstChild.IsComplete AND SecondChild.IsComplete
                AND (FirstChild.Result = E_Result.Passed) AND (SecondChild.Result = E_Result.Passed);
            FCompletedRuns := FCompletedRuns + 1;
            CheckReservations();
            CheckEventStream();
            IF FCompletedRuns = RequiredRuns THEN
                FStep := Finish;
            ELSE
                FStep := ResetRequested;
            END_IF;
        END_IF;
END_CASE;
END_METHOD

END_FUNCTION_BLOCK

// ---- SelfTests/TestCases/TestSuite_RunControlLifecycle/Helper/RunControlIntegrationSubject.TcPOU
{region 'Documentation'}
(*!
<summary>Local real root, Orchestrator, Suite and two Test Cases with one isolated publisher.</summary>
<description>
BindPublisher wires each producer before Initialize. Production lifecycle, scheduling and
reservation handling remain inherited. Configure initializes the hierarchy once; lifecycle
Reset does not rebuild it. Observation accessors expose the actual children, not mirrored state.
</description>
*)
{endregion}
FUNCTION_BLOCK RunControlIntegrationSubject EXTENDS RunControlBase
VAR
    FSuite : SuiteIntegrationSubject;
    FTestSuites : ARRAY[3..4] OF I_TestSuite;
    FRealOrchestrator : OrchestratorProbe;
    FConfigureCount : UINT;
END_VAR

SUPER^(ControlData := ControlData);

{region 'Documentation'}
(*!
<summary>Binds the complete local hierarchy before first use without changing the global publisher.</summary>
*)
{endregion}
METHOD PUBLIC BindPublisher
VAR_INPUT
    Publisher : I_EventPublisher; //! Nonzero isolated event publisher retained before subject initialization; keep it alive through all subject use.
END_VAR
FEventPublisher := Publisher;
FRealOrchestrator.BindPublisher(Publisher := Publisher);
FOrchestrator := FRealOrchestrator;
FSuite.BindPublisher(Publisher := Publisher);
FConfigureCount := 0;
END_METHOD

{region 'Documentation'}
(*!
<summary>Reports the Suite's observation of exactly one call per concrete Test Case.</summary>
*)
{endregion}
{attribute 'monitoring' := 'call'}
PROPERTY PUBLIC ChildCallsMatch : BOOL //! Reports the Suite's observation of exactly one call per concrete Test Case.
GET
ChildCallsMatch := FSuite.ChildCallsMatch;
END_GET
END_PROPERTY

{region 'Documentation'}
(*!
<summary>Confirms both owner configurations ran once across lifecycle Reset/repeat.</summary>
*)
{endregion}
{attribute 'monitoring' := 'call'}
PROPERTY PUBLIC ConfigurationUnchanged : BOOL //! Confirms both owner configurations ran once across lifecycle Reset/repeat.
GET
ConfigurationUnchanged := (FConfigureCount = 1) AND (FSuite.ConfigureCount = 1);
END_GET
END_PROPERTY

{region 'Documentation'}
(*!
<summary>Registers one real Suite; normal configuration defaults include the completion delay.</summary>
*)
{endregion}
METHOD PROTECTED Configure
VAR_IN_OUT
    // SA0167: Borrowed owner builder; no temporary instance is created.
    {attribute 'analysis' := '-167'}
    Builder : RunControlConfigurationBuilder; //! Borrowed owner configuration builder used only during this Configure call; register this owner's concrete children.
END_VAR
VAR
    Config : ST_TestSuiteConfig;
END_VAR
FConfigureCount := FConfigureCount + 1;
Builder.Initialize(Mode := E_OrchestrationMode.Serial,
    TestSuites := FTestSuites);
FSuite.Initialize(Parent := THIS^,
    SuiteName := 'Suite',
    Config := Config);
Builder.Register(TestSuite := FSuite);
END_METHOD

{region 'Documentation'}
(*!
<summary>Provides the actual Suite child by its registered index for integration observations.</summary>
*)
{endregion}
METHOD PUBLIC GetTestCase : I_TestCase //! Typed child interface at the original array index; zero when no entry is available.
VAR_INPUT
    Index : DINT; //! Original occupied child-array index, rather than an ordinal position.
END_VAR
GetTestCase := FSuite.GetTestCase(Index := Index);
END_METHOD

{region 'Documentation'}
(*!
<summary>Returns the registered Suite for its original array index.</summary>
*)
{endregion}
METHOD PUBLIC GetTestSuite : I_TestSuite //! Typed Suite interface at the original array index; zero when no entry is available.
VAR_INPUT
    Index : DINT; //! Original occupied child-array index, rather than an ordinal position.
END_VAR
GetTestSuite := 0;
IF (ChildCount = 0) OR (Index <> ChildArrayLowerBound) THEN
    RETURN;
END_IF;
GetTestSuite := FTestSuites[Index];
END_METHOD

{region 'Documentation'}
(*!
<summary>Calls the owned real Suite once per root cycle, including Completed.</summary>
*)
{endregion}
METHOD PROTECTED ProcessTestSuites
FSuite();
END_METHOD

{region 'Documentation'}
(*!
<summary>First registered Test Case array index in the real Suite.</summary>
*)
{endregion}
{attribute 'monitoring' := 'call'}
PROPERTY PUBLIC TestCaseLowerBound : DINT //! First registered Test Case array index in the real Suite.
GET
TestCaseLowerBound := FSuite.ChildArrayLowerBound;
END_GET
END_PROPERTY

END_FUNCTION_BLOCK

// ---- SelfTests/TestCases/TestSuite_RunControlLifecycle/Test_RunControlExceptionalLifecycle.TcPOU
{region 'Documentation'}
(*!
<summary>Exercises Root error and Abort paths through controlled child/helper observations.</summary>
<description>

Scenario ownership

Each instance runs one selected scenario. Production root sequencing, timers, result handling
and publication stay unchanged. The local helper supplies observations, never child scheduling.
Only the isolated subject writes to the local capture; checking Assertions use the normal publisher.

Script and call order

RunStep arranges one cycle, calls the subject once, then checks the expected owner response.
FNextStep is accepted only after checking Assertions ran. Child snapshots are applied by the
subject's ProcessTestSuites, so child errors affect the result in that call and the next Sequencer call.

Timeout and recovery

Timeout scenarios withhold completion for the real configured deadline. Waiting
repeats a checkpoint, not subject calls within a cycle. The outer Test Case timeout bounds a
missing transition. An independent scheduled-task stopwatch checks that deadlines are neither early nor restarted
on Abort-to-error escalation. This checks lifecycle timing, not physical clock calibration.
Completed calls continue child processing, including late child completion after root timeout.
A recorded interface-call boundary verifies that the root leaves child requests and resource
release to its selected helper rather than adding direct cleanup calls. The controlled helper
itself does not model reservations; real resource release belongs to composition integration.
Every scenario ends with a successful lifecycle Reset without replacing bindings or configuration.
</description>
*)
{endregion}
FUNCTION_BLOCK Test_RunControlExceptionalLifecycle EXTENDS TestCaseBase
VAR_INPUT
    Scenario : E_RunControlLifecycleScenario := E_RunControlLifecycleScenario.ResetError; //! Fixed scenario selection supplied by the containing Suite on every call.
END_VAR
VAR
    FControl : ST_RunControl;
    FDeadlineTimer : Stopwatch;
    FCompletedSequence : UDINT;
    FSubject : RunControlLifecycleProbe;
    FHelper : SuiteOrchestratorDouble;
    FCapture : EventBuffer;
    FEvents : ARRAY[1..CaptureLength] OF ST_Event;
    FCaptureFifo : ST_FifoStatus;
    FCaptureStatus : ST_EventBufferStatus;
    FFirstChild : ST_OrchestrationObservation;
    FSecondChild : ST_OrchestrationObservation;
    FStep : INT;
    FNextStep : INT;
    FStepChecked : BOOL;
    FSubjectCallCount : UINT;
    FExpectedTimeout : BOOL;
    FExpectedResetTimeout : BOOL;
    FExpectedAbortTimeout : BOOL;
    FStatePath : AssertTrue;
    FStatePathMatches : BOOL := TRUE;
    FTaskMapping : AssertTrue;
    FTaskMappingMatches : BOOL := TRUE;
    FResultStatus : AssertTrue;
    FResultStatusMatches : BOOL := TRUE;
    FTimeoutFlags : AssertTrue;
    FTimeoutFlagsMatches : BOOL := TRUE;
    FChildCalls : AssertTrue;
    FChildCallsMatches : BOOL := TRUE;
    FEventEvidence : AssertTrue;
    FEventEvidenceMatches : BOOL := TRUE;
    FDeadline : AssertTrue;
    FDeadlineMatches : BOOL := TRUE;
    FDelegation : AssertTrue;
    FDelegationMatches : BOOL := TRUE;
    FRecovery : AssertTrue;
    FRecoveryMatches : BOOL := TRUE;
END_VAR
VAR CONSTANT
    CaptureLength : UINT := 64;
    ShortTimeout : TIME := T#50ms;
    Setup : INT := 0;
    ObserveInitialReset : INT := 1;
    InitialResetResponse : INT := 2;
    HoldResetError : INT := 3;
    FinishFailedReset : INT := 4;
    StartExecution : INT := 5;
    ReachRunning : INT := 6;
    ApplyStimulus : INT := 7;
    ObserveChildError : INT := 8;
    ObserveAbortResponse : INT := 9;
    FinishChildren : INT := 10;
    FinishHelper : INT := 11;
    CheckCompleted : INT := 12;
    HoldCompleted : INT := 13;
    LateChildrenFinish : INT := 14;
    RecoveryReset : INT := 15;
    RecoveryReady : INT := 16;
    Done : INT := 17;
    AwaitEscalatedAbortTimeout : INT := 18;
END_VAR

SUPER^();

{region 'Documentation'}
(*!
<summary>Contributes only the checking Assertions, not the intentionally controlled subject results.</summary>
*)
{endregion}
METHOD PROTECTED AggregateResults
VAR_INPUT
    Aggregator : I_ResultAggregator; //! Borrowed result sink owned by the outer Test Case; add this test's checking Assertions without resetting or retaining the sink.
END_VAR
Aggregator.AddProvider(Provider := FStatePath);
Aggregator.AddProvider(Provider := FTaskMapping);
Aggregator.AddProvider(Provider := FResultStatus);
Aggregator.AddProvider(Provider := FTimeoutFlags);
Aggregator.AddProvider(Provider := FChildCalls);
Aggregator.AddProvider(Provider := FEventEvidence);
Aggregator.AddProvider(Provider := FRecovery);
Aggregator.AddProvider(Provider := FDeadline);
Aggregator.AddProvider(Provider := FDelegation);
END_METHOD

{region 'Documentation'}
(*!
<summary>Checks exceptional finalization and diagnostics; failed Reset must have no Abort transition.</summary>
*)
{endregion}
METHOD PRIVATE CheckEventEvidence
VAR
    Index : UINT;
    DiagnosticCount : UINT;
    AbortTransitionCount : UINT;
    ResultCount : UINT;
    AggregationCount : UINT;
    CompletedCount : UINT;
    ResultSequence : UDINT;
    AggregationSequence : UDINT;
    CompletedSequence : UDINT;
    ExpectedResult : E_Result := E_Result.Error;
    PayloadMatches : BOOL := TRUE;
END_VAR
IF Scenario = E_RunControlLifecycleScenario.Abort THEN
    ExpectedResult := E_Result.Abort;
END_IF;
FOR Index := 1 TO CaptureLength DO
    IF (FEvents[Index].SequenceId = 0) OR (FEvents[Index].Name <> FSubject.Name) THEN
        CONTINUE;
    END_IF;
    CASE FEvents[Index].EventType OF
        E_EventType.Result:
            ResultCount := ResultCount + 1;
            ResultSequence := FEvents[Index].SequenceId;
            PayloadMatches := PayloadMatches
                AND (FEvents[Index].OwnerScope = E_OwnerScope.RunControl)
                AND (FEvents[Index].State = E_State.Completing)
                AND (FEvents[Index].Result = ExpectedResult);
        E_EventType.Aggregation:
            AggregationCount := AggregationCount + 1;
            AggregationSequence := FEvents[Index].SequenceId;
            PayloadMatches := PayloadMatches
                AND (FEvents[Index].OwnerScope = E_OwnerScope.RunControl)
                AND (FEvents[Index].State = E_State.Completing)
                AND (FEvents[Index].Result = ExpectedResult);
        E_EventType.StateTransition:
            IF FEvents[Index].State = E_State.Completed THEN
                CompletedCount := CompletedCount + 1;
                CompletedSequence := FEvents[Index].SequenceId;
            END_IF;
    END_CASE;
    IF (FEvents[Index].EventType = E_EventType.Framework)
        AND (FEvents[Index].Severity = E_EventSeverity.Error) THEN
        DiagnosticCount := DiagnosticCount + 1;
    END_IF;
    IF (FEvents[Index].EventType = E_EventType.StateTransition)
        AND ((FEvents[Index].State = E_State.Aborting)
            OR (FEvents[Index].State = E_State.AbortingFromError)) THEN
        AbortTransitionCount := AbortTransitionCount + 1;
    END_IF;
END_FOR;
IF Scenario = E_RunControlLifecycleScenario.Abort THEN
    FEventEvidenceMatches := DiagnosticCount = 0;
ELSIF (Scenario = E_RunControlLifecycleScenario.ResetErrorTimeout)
    OR (Scenario = E_RunControlLifecycleScenario.AbortErrorTimeout) THEN
    FEventEvidenceMatches := DiagnosticCount = 2;
ELSE
    FEventEvidenceMatches := DiagnosticCount = 1;
END_IF;
IF (Scenario = E_RunControlLifecycleScenario.ResetError) OR (Scenario = E_RunControlLifecycleScenario.ResetTimeout)
    OR (Scenario = E_RunControlLifecycleScenario.ResetErrorTimeout) THEN
    FEventEvidenceMatches := FEventEvidenceMatches AND (AbortTransitionCount = 0);
ELSE
    FEventEvidenceMatches := FEventEvidenceMatches AND (AbortTransitionCount > 0);
END_IF;
FEventEvidenceMatches := FEventEvidenceMatches AND PayloadMatches
    AND (ResultCount = 1) AND (AggregationCount = 1) AND (CompletedCount = 1)
    AND (ResultSequence < AggregationSequence) AND (AggregationSequence < CompletedSequence)
    AND (FCaptureStatus.LostEventCount = 0);
END_METHOD

{region 'Documentation'}
(*!
<summary>Initializes the checking Assertions; the scenario explicitly initializes its isolated subject.</summary>
*)
{endregion}
METHOD PROTECTED Configure
FPreparationStateCount := 0;
FTestStateCount := 1;
FStatePath.Initialize(Parent := THIS^,
    AssertionName := 'StatePath');
FTaskMapping.Initialize(Parent := THIS^,
    AssertionName := 'TaskMapping');
FResultStatus.Initialize(Parent := THIS^,
    AssertionName := 'ResultStatus');
FTimeoutFlags.Initialize(Parent := THIS^,
    AssertionName := 'TimeoutFlags');
FChildCalls.Initialize(Parent := THIS^,
    AssertionName := 'ChildCalls');
FEventEvidence.Initialize(Parent := THIS^,
    AssertionName := 'EventEvidence');
FRecovery.Initialize(Parent := THIS^,
    AssertionName := 'Recovery');
FDeadline.Initialize(Parent := THIS^,
    AssertionName := 'Deadline');
FDelegation.Initialize(Parent := THIS^,
    AssertionName := 'Delegation');
END_METHOD

{region 'Documentation'}
(*!
<summary>No asynchronous test resource remains to stop.</summary>
*)
{endregion}
METHOD PROTECTED ProcessAbort
VAR_INPUT
    Enable : BOOL; //! Phase permission supplied by the owning Test Case; FALSE does not authorize progression, while observation may continue.
END_VAR
IF Enable THEN
    CompleteAbort();
END_IF;
END_METHOD

{region 'Documentation'}
(*!
<summary>Checks every subject cycle before advancing, retaining failures across waiting and recovery.</summary>
*)
{endregion}
METHOD PROTECTED ProcessAssertions
VAR_INPUT
    Enable : BOOL; //! Phase permission supplied by the owning Test Case; FALSE does not authorize progression, while observation may continue.
END_VAR
FStatePath(Enable := Enable,
    State := State,
    IN := FStatePathMatches);
FTaskMapping(Enable := Enable,
    State := State,
    IN := FTaskMappingMatches);
FResultStatus(Enable := Enable,
    State := State,
    IN := FResultStatusMatches);
FTimeoutFlags(Enable := Enable,
    State := State,
    IN := FTimeoutFlagsMatches);
FChildCalls(Enable := Enable,
    State := State,
    IN := FChildCallsMatches);
FEventEvidence(Enable := Enable,
    State := State,
    IN := FEventEvidenceMatches);
FRecovery(Enable := Enable,
    State := State,
    IN := FRecoveryMatches);
FDeadline(Enable := Enable,
    State := State,
    IN := FDeadlineMatches);
FDelegation(Enable := Enable,
    State := State,
    IN := FDelegationMatches);
IF Enable THEN
    FStepChecked := TRUE;
END_IF;
END_METHOD

{region 'Documentation'}
(*!
<summary>No resource Preparation is required for this controlled owner scenario.</summary>
*)
{endregion}
METHOD PROTECTED ProcessPreparations
VAR_INPUT
    // SA0033: Required override; the scenario has no Preparation phase.
    {attribute 'analysis' := '-33'}
    Enable : BOOL; //! Phase permission supplied by the owning Test Case; FALSE does not authorize progression, while observation may continue.
END_VAR
END_METHOD

{region 'Documentation'}
(*!
<summary>Restarts the test script and clears checking Assertions; subject setup belongs to the next test attempt.</summary>
*)
{endregion}
METHOD PROTECTED ProcessReset
FStep := Setup;
FNextStep := Setup;
FStepChecked := FALSE;
FSubjectCallCount := 0;
FExpectedTimeout := FALSE;
FExpectedResetTimeout := FALSE;
FExpectedAbortTimeout := FALSE;
FStatePathMatches := TRUE;
FTaskMappingMatches := TRUE;
FResultStatusMatches := TRUE;
FTimeoutFlagsMatches := TRUE;
FChildCallsMatches := TRUE;
FEventEvidenceMatches := TRUE;
FRecoveryMatches := TRUE;
FStatePath.Reset();
FTaskMapping.Reset();
FResultStatus.Reset();
FTimeoutFlags.Reset();
FChildCalls.Reset();
FEventEvidence.Reset();
FRecovery.Reset();
FDeadline.Reset();
FDelegation.Reset();
FDeadlineMatches := TRUE;
FDelegationMatches := TRUE;
FDeadlineTimer.Reset();
FCompletedSequence := 0;
CompleteReset();
END_METHOD

{region 'Documentation'}
(*!
<summary>Advances the explicit test script with at most one subject FB call per active PLC cycle.</summary>
*)
{endregion}
METHOD PROTECTED ProcessTests
VAR_INPUT
    Enable : BOOL; //! Phase permission supplied by the owning Test Case; FALSE does not authorize progression, while observation may continue.
END_VAR
IF NOT Enable THEN
    RETURN;
END_IF;
IF FStepChecked THEN
    FStep := FNextStep;
    FStepChecked := FALSE;
END_IF;
IF FStep = Done THEN
    CompleteTests();
    RETURN;
END_IF;
RunStep();
END_METHOD

{region 'Documentation'}
(*!
<summary>Arranges one error-path checkpoint and checks the real root; timeout waits use further PLC cycles.</summary>
*)
{endregion}
METHOD PRIVATE RunStep
VAR
    Config : ST_RunConfig;
    Snapshot : ST_RunControlStatus;
    ExpectedState : E_State;
    ExpectedTask : E_OrchestratorTask;
    ExpectedResult : E_Result;
    FinalResult : E_Result;
    WaitForTimeout : BOOL;
    WaitingState : E_State;
    WaitingTask : E_OrchestratorTask;
    WaitingResult : E_Result := E_Result.NotEvaluated;
    FirstCalls : ST_OrchestrationCalls;
    LastCalls : ST_OrchestrationCalls;
END_VAR
FDeadlineTimer.Update();
FNextStep := FStep + 1;
ExpectedResult := E_Result.NotEvaluated;
ExpectedTask := E_OrchestratorTask.Idle;
FinalResult := E_Result.Error;
IF Scenario = E_RunControlLifecycleScenario.Abort THEN
    FinalResult := E_Result.Abort;
END_IF;

CASE FStep OF
    Setup:
        CASE Scenario OF
            E_RunControlLifecycleScenario.ResetTimeout, E_RunControlLifecycleScenario.ResetErrorTimeout:
                Config.ResetTimeout := ShortTimeout;
            E_RunControlLifecycleScenario.ExecutionTimeout:
                Config.Timeout := ShortTimeout;
            E_RunControlLifecycleScenario.AbortTimeout, E_RunControlLifecycleScenario.AbortErrorTimeout:
                Config.AbortTimeout := ShortTimeout;
        ELSE
            // Other scenarios use the ordinary positive deadlines.
        END_CASE;
        Config.CompletionDelay := T#0ms;
        IF NOT FCapture.Initialize(Buffer := FEvents,
            FifoControl := FCaptureFifo,
            Status := FCaptureStatus) THEN
            Error(Message := 'Exceptional root capture could not be initialized.');
            RETURN;
        END_IF;
        FHelper.BeginScenario();
        FSubject.Bind(Publisher := FCapture,
            Helper := FHelper,
            Config := Config);
        IF NOT FSubject.Initialize(Name := 'ExceptionalSubject',
            EventBuffer := FCapture) THEN
            Error(Message := 'Exceptional root subject could not be initialized.');
            RETURN;
        END_IF;
        FDeadlineTimer.Start();
        FFirstChild.State := E_State.Reset;
        FFirstChild.Result := E_Result.NotEvaluated;
        FFirstChild.Ready := FALSE;
        FFirstChild.Complete := FALSE;
        FSecondChild := FFirstChild;
        ExpectedState := E_State.Reset;
        ExpectedTask := E_OrchestratorTask.Reset;

    ObserveInitialReset:
        FFirstChild.State := E_State.Reset;
        FSecondChild := FFirstChild;
        ExpectedState := E_State.Reset;
        ExpectedTask := E_OrchestratorTask.Reset;

    InitialResetResponse:
        CASE Scenario OF
            E_RunControlLifecycleScenario.ResetError, E_RunControlLifecycleScenario.ResetErrorTimeout:
                FHelper.SetObservation(Ready := FALSE,
                    Result := E_Result.Error);
                FFirstChild.State := E_State.Completed;
                FFirstChild.Result := E_Result.Error;
                FFirstChild.Complete := TRUE;
                ExpectedState := E_State.Reset;
                ExpectedResult := E_Result.Error;
                ExpectedTask := E_OrchestratorTask.Reset;
                FNextStep := HoldResetError;

            E_RunControlLifecycleScenario.ResetTimeout:
                WaitForTimeout := TRUE;
                WaitingState := E_State.Reset;
                WaitingTask := E_OrchestratorTask.Reset;
                ExpectedState := E_State.Completing;
                ExpectedResult := E_Result.Error;
                FNextStep := CheckCompleted;
        ELSE
            FHelper.SetObservation(Ready := TRUE,
                ResetFinished := TRUE);
            FFirstChild.State := E_State.Idle;
            FFirstChild.Ready := TRUE;
            FSecondChild := FFirstChild;
            ExpectedState := E_State.Idle;
            FNextStep := StartExecution;
        END_CASE;

    HoldResetError:
        // Another Reset request must not clear the held error or abandon the unfinished child.
        FSubject.RequestReset();
        ExpectedState := E_State.Reset;
        ExpectedResult := E_Result.Error;
        ExpectedTask := E_OrchestratorTask.Reset;

    FinishFailedReset:
        ExpectedState := E_State.Completing;
        ExpectedResult := E_Result.Error;
        FNextStep := CheckCompleted;
        IF Scenario = E_RunControlLifecycleScenario.ResetErrorTimeout THEN
            WaitForTimeout := TRUE;
            WaitingState := E_State.Reset;
            WaitingTask := E_OrchestratorTask.Reset;
            WaitingResult := E_Result.Error;
        ELSE
            FHelper.SetObservation(Ready := FALSE,
                Result := E_Result.Error,
                ResetFinished := TRUE);
            FSecondChild.State := E_State.Idle;
            FSecondChild.Ready := TRUE;
        END_IF;

    StartExecution:
        FDeadlineTimer.Start();
        FSubject.RequestStart();
        FFirstChild.State := E_State.Running;
        FFirstChild.Ready := FALSE;
        ExpectedState := E_State.Starting;
        ExpectedTask := E_OrchestratorTask.Execution;

    ReachRunning:
        FHelper.SetObservation(Ready := FALSE);
        ExpectedState := E_State.Running;
        ExpectedTask := E_OrchestratorTask.Execution;

    ApplyStimulus:
        CASE Scenario OF
            E_RunControlLifecycleScenario.ChildError, E_RunControlLifecycleScenario.UnexpectedChildAbort:
                FFirstChild.State := E_State.Completed;
                FFirstChild.Complete := TRUE;
                IF Scenario = E_RunControlLifecycleScenario.ChildError THEN
                    FFirstChild.Result := E_Result.Error;
                ELSE
                    FFirstChild.Result := E_Result.Abort;
                END_IF;
                ExpectedState := E_State.Running;
                ExpectedResult := E_Result.Error;
                ExpectedTask := E_OrchestratorTask.Execution;
                FNextStep := ObserveChildError;

            E_RunControlLifecycleScenario.ExecutionError:
                FHelper.SetObservation(Ready := FALSE,
                    Result := E_Result.Error);
                ExpectedState := E_State.AbortingFromError;
                ExpectedResult := E_Result.Error;
                ExpectedTask := E_OrchestratorTask.Abort;
                FNextStep := FinishChildren;

            E_RunControlLifecycleScenario.ExecutionTimeout:
                WaitForTimeout := TRUE;
                WaitingState := E_State.Running;
                WaitingTask := E_OrchestratorTask.Execution;
                ExpectedState := E_State.AbortingFromError;
                ExpectedResult := E_Result.Error;
                ExpectedTask := E_OrchestratorTask.Abort;
                FNextStep := FinishChildren;

            E_RunControlLifecycleScenario.Abort, E_RunControlLifecycleScenario.AbortError,
                E_RunControlLifecycleScenario.AbortTimeout, E_RunControlLifecycleScenario.AbortErrorTimeout:
                FDeadlineTimer.Start();
                FSubject.RequestAbort();
                FFirstChild.State := E_State.Aborting;
                FFirstChild.Result := E_Result.Abort;
                ExpectedState := E_State.Aborting;
                ExpectedResult := E_Result.Abort;
                ExpectedTask := E_OrchestratorTask.Abort;
                FNextStep := ObserveAbortResponse;
        ELSE
            Error(Message := 'Unsupported execution stimulus.');
            RETURN;
        END_CASE;

    ObserveChildError:
        ExpectedState := E_State.AbortingFromError;
        ExpectedResult := E_Result.Error;
        ExpectedTask := E_OrchestratorTask.Abort;
        FNextStep := FinishChildren;

    ObserveAbortResponse:
        CASE Scenario OF
            E_RunControlLifecycleScenario.Abort:
                ExpectedState := E_State.Aborting;
                ExpectedResult := E_Result.Abort;
                ExpectedTask := E_OrchestratorTask.Abort;
                FNextStep := FinishChildren;
            E_RunControlLifecycleScenario.AbortError:
                FHelper.SetObservation(Ready := FALSE,
                    Result := E_Result.Error);
                ExpectedState := E_State.AbortingFromError;
                ExpectedResult := E_Result.Error;
                ExpectedTask := E_OrchestratorTask.Abort;
                FNextStep := FinishChildren;
            E_RunControlLifecycleScenario.AbortErrorTimeout:
                ExpectedTask := E_OrchestratorTask.Abort;
                IF FDeadlineTimer.ElapsedLTime < TIME_TO_LTIME(ShortTimeout) / 2 THEN
                    ExpectedState := E_State.Aborting;
                    ExpectedResult := E_Result.Abort;
                    FNextStep := ObserveAbortResponse;
                ELSE
                    FHelper.SetObservation(Ready := FALSE,
                        Result := E_Result.Error);
                    ExpectedState := E_State.AbortingFromError;
                    ExpectedResult := E_Result.Error;
                    FNextStep := AwaitEscalatedAbortTimeout;
                END_IF;
            E_RunControlLifecycleScenario.AbortTimeout:
                WaitForTimeout := TRUE;
                WaitingState := E_State.Aborting;
                WaitingResult := E_Result.Abort;
                WaitingTask := E_OrchestratorTask.Abort;
                ExpectedState := E_State.Completing;
                ExpectedResult := E_Result.Error;
                ExpectedTask := E_OrchestratorTask.Abort;
                FNextStep := CheckCompleted;
        ELSE
            Error(Message := 'Unsupported Abort observation.');
            RETURN;
        END_CASE;

    AwaitEscalatedAbortTimeout:
        WaitForTimeout := TRUE;
        WaitingState := E_State.AbortingFromError;
        WaitingResult := E_Result.Error;
        WaitingTask := E_OrchestratorTask.Abort;
        ExpectedState := E_State.Completing;
        ExpectedResult := E_Result.Error;
        ExpectedTask := E_OrchestratorTask.Abort;
        FNextStep := CheckCompleted;

    FinishChildren:
        FFirstChild.State := E_State.Completed;
        FFirstChild.Ready := FALSE;
        FFirstChild.Complete := TRUE;
        IF Scenario <> E_RunControlLifecycleScenario.ChildError THEN
            FFirstChild.Result := E_Result.Abort;
        END_IF;
        ExpectedState := E_State.AbortingFromError;
        IF Scenario = E_RunControlLifecycleScenario.Abort THEN
            ExpectedState := E_State.Aborting;
        END_IF;
        ExpectedResult := FinalResult;
        ExpectedTask := E_OrchestratorTask.Abort;

    FinishHelper:
        FHelper.SetObservation(Ready := FALSE,
            Result := FHelper.Result,
            AbortFinished := TRUE);
        ExpectedState := E_State.Completing;
        ExpectedResult := FinalResult;
        ExpectedTask := E_OrchestratorTask.Abort;

    CheckCompleted, HoldCompleted:
        ExpectedState := E_State.Completed;
        ExpectedResult := FinalResult;

    LateChildrenFinish:
        IF NOT FFirstChild.Complete THEN
            FFirstChild.State := E_State.Completed;
            FFirstChild.Result := E_Result.Error;
            FFirstChild.Complete := TRUE;
            FFirstChild.Ready := FALSE;
        END_IF;
        FSecondChild.State := E_State.Idle;
        FSecondChild.Result := E_Result.NotEvaluated;
        FSecondChild.Complete := FALSE;
        FSecondChild.Ready := TRUE;
        ExpectedState := E_State.Completed;
        ExpectedResult := FinalResult;

    RecoveryReset:
        FHelper.SetObservation(Ready := FALSE);
        FSubject.RequestReset();
        FFirstChild.State := E_State.Reset;
        FFirstChild.Result := E_Result.NotEvaluated;
        FFirstChild.Complete := FALSE;
        FFirstChild.Ready := FALSE;
        FSecondChild := FFirstChild;
        FExpectedTimeout := FALSE;
        FExpectedResetTimeout := FALSE;
        FExpectedAbortTimeout := FALSE;
        ExpectedState := E_State.Reset;
        ExpectedTask := E_OrchestratorTask.Reset;

    RecoveryReady:
        FHelper.SetObservation(Ready := TRUE,
            ResetFinished := TRUE);
        FFirstChild.State := E_State.Idle;
        FFirstChild.Ready := TRUE;
        FSecondChild := FFirstChild;
        ExpectedState := E_State.Idle;
ELSE
    Error(Message := 'Unexpected exceptional root test step.');
    RETURN;
END_CASE;

FSubject.SetChildObservations(FirstChild := FFirstChild,
    SecondChild := FSecondChild);
FSubject(ControlData := FControl);
FSubjectCallCount := FSubjectCallCount + 1;
Snapshot := FSubject.Status;

IF WaitForTimeout THEN
    IF FSubject.State = WaitingState THEN
        ExpectedState := WaitingState;
        ExpectedTask := WaitingTask;
        ExpectedResult := WaitingResult;
        FNextStep := FStep;
        FDeadlineMatches := FDeadlineTimer.IsValid
            AND (FDeadlineTimer.ElapsedLTime < TIME_TO_LTIME(ShortTimeout));
    ELSE
        FDeadlineMatches := FDeadlineTimer.IsValid
            AND (FDeadlineTimer.ElapsedLTime >= TIME_TO_LTIME(ShortTimeout));
        CASE Scenario OF
            E_RunControlLifecycleScenario.ResetTimeout, E_RunControlLifecycleScenario.ResetErrorTimeout:
                FExpectedResetTimeout := TRUE;
            E_RunControlLifecycleScenario.ExecutionTimeout:
                FExpectedTimeout := TRUE;
            E_RunControlLifecycleScenario.AbortTimeout, E_RunControlLifecycleScenario.AbortErrorTimeout:
                FExpectedAbortTimeout := TRUE;
        ELSE
            Error(Message := 'Unexpected timeout-wait scenario.');
            RETURN;
        END_CASE;
    END_IF;
END_IF;

FStatePathMatches := (FSubject.State = ExpectedState)
    AND (Snapshot.Execution.State = ExpectedState)
    AND (FControl.Status.Execution.State = ExpectedState)
    AND (FControl.Name = FSubject.Name);
FTaskMappingMatches := FHelper.CurrentTask = ExpectedTask;
FResultStatusMatches := (FSubject.Result = ExpectedResult)
    AND (Snapshot.Execution.Result = ExpectedResult)
    AND (FControl.Status.Execution.Result = ExpectedResult)
    AND (FSubject.HasError = (ExpectedResult = E_Result.Error))
    AND (Snapshot.Execution.Error = (ExpectedResult = E_Result.Error))
    AND (FSubject.IsComplete = (ExpectedState = E_State.Completed))
    AND (Snapshot.Execution.Completed = (ExpectedState = E_State.Completed));
FTimeoutFlagsMatches := (FSubject.HasTimeout = FExpectedTimeout)
    AND (FSubject.HasResetTimeout = FExpectedResetTimeout)
    AND (FSubject.HasAbortTimeout = FExpectedAbortTimeout);
FChildCallsMatches := (FHelper.ExecuteCount = FSubjectCallCount)
    AND (FSubject.ChildCallCount = FSubjectCallCount)
    AND FSubject.ChildBodyCallsMatch;

FirstCalls := FSubject.GetChildCalls(Index := FSubject.ChildArrayLowerBound);
LastCalls := FSubject.GetChildCalls(Index := FSubject.ChildArrayLowerBound + UINT_TO_DINT(FSubject.ChildCount) - 1);
FDelegationMatches := (FirstCalls.StartCount = 0) AND (LastCalls.StartCount = 0)
    AND (FirstCalls.ResetCount = 0) AND (LastCalls.ResetCount = 0)
    AND (FirstCalls.AbortCount = 0) AND (LastCalls.AbortCount = 0)
    AND (FirstCalls.ExecutionReservationCount = 0) AND (LastCalls.ExecutionReservationCount = 0)
    AND (FirstCalls.ResetReservationCount = 0) AND (LastCalls.ResetReservationCount = 0)
    AND (FirstCalls.FreeCount = 0) AND (LastCalls.FreeCount = 0);
IF (FStep = CheckCompleted) OR (FStep = HoldCompleted) OR (FStep = LateChildrenFinish) THEN
    CheckEventEvidence();
    IF FStep = CheckCompleted THEN
        FCompletedSequence := FCaptureStatus.SequenceId;
    ELSE
        FEventEvidenceMatches := FEventEvidenceMatches AND (FCaptureStatus.SequenceId = FCompletedSequence);
    END_IF;
END_IF;
IF FStep = LateChildrenFinish THEN
    FChildCallsMatches := FChildCallsMatches
        AND (Snapshot.SuiteCountCompleted = 1) AND (Snapshot.SuiteCountIdle = 1);
END_IF;
IF FStep = RecoveryReady THEN
    FRecoveryMatches := FSubject.IsReady AND Snapshot.Execution.Ready
        AND (FSubject.Result = E_Result.NotEvaluated)
        AND (FHelper.InitializeCount = 1) AND (FSubject.ConfigureCount = 1)
        AND (FCapture.ReservedEntryCount = 0)
        AND (FCaptureStatus.LostEventCount = 0);
END_IF;
END_METHOD

END_FUNCTION_BLOCK

// ---- SelfTests/TestCases/TestSuite_RunControlLifecycle/Test_RunControlCompletion.TcPOU
{region 'Documentation'}
(*!
<summary>Checks root completion timing, frozen event payloads and live child observations.</summary>
<description>

Ownership and steps

Each instance selects one fixed scenario. A real RunControlBase uses a controlled helper
and two Suite observations, with a private Event Buffer. RunStep arranges one subject call;
checking Assertions consume the observations before the next step is accepted.

Clock observation

ZeroDelay and DefaultDelay use the unchanged production clock. The independent stopwatch
starts in the entry cycle of Completing. Completed must occur on a later call, never before
the configured interval. InvalidTime overrides only the agreed validity observation after
final events exist; it does not change task time, elapsed values or transition logic.

Publication versus status

The entry Result and Aggregation are checked and retained. Subsequent calls verify every
event field and prohibit republication. LateResetChildren leaves a child resetting when
the root times out; its later completion changes live counters without rewriting the log.
Every case holds Completed for further calls and then verifies ordinary Reset recovery.
</description>
*)
{endregion}
FUNCTION_BLOCK Test_RunControlCompletion EXTENDS TestCaseBase
VAR_INPUT
    Scenario : E_RunControlCompletionScenario := E_RunControlCompletionScenario.DefaultDelay; //! Completion scenario selected by the containing Suite and held fixed during this instance.
END_VAR
VAR
    FSubject : RunControlLifecycleProbe;
    FHelper : SuiteOrchestratorDouble;
    FControl : ST_RunControl;
    FCapture : EventBuffer;
    FEvents : ARRAY[1..CaptureLength] OF ST_Event;
    FCaptureFifo : ST_FifoStatus;
    FCaptureStatus : ST_EventBufferStatus;
    FFirstChild : ST_OrchestrationObservation;
    FSecondChild : ST_OrchestrationObservation;
    FDelayClock : Stopwatch;
    FDelay : TIME;
    FExpectedResult : E_Result;
    FPublishedResult : ST_Event;
    FPublishedAggregation : ST_Event;
    FFinalRuntime : TIME;
    FStep : INT;
    FNextStep : INT;
    FStepChecked : BOOL;
    FCallCount : UINT;
    FEntryCall : UINT;
    FHoldCalls : UINT;
    FStatePath : AssertTrue;
    FStatePathMatches : BOOL := TRUE;
    FTiming : AssertTrue;
    FTimingMatches : BOOL := TRUE;
    FFinalEvents : AssertTrue;
    FFinalEventsMatches : BOOL := TRUE;
    FPublishedPayload : AssertTrue;
    FPublishedPayloadMatches : BOOL := TRUE;
    FLiveStatus : AssertTrue;
    FLiveStatusMatches : BOOL := TRUE;
    FDiagnostics : AssertTrue;
    FDiagnosticsMatches : BOOL := TRUE;
    FChildCalls : AssertTrue;
    FChildCallsMatches : BOOL := TRUE;
    FRecovery : AssertTrue;
    FRecoveryMatches : BOOL := TRUE;
END_VAR
VAR CONSTANT
    CaptureLength : UINT := 64;
    DefaultDelay : TIME := T#100ms;
    ResetDeadline : TIME := T#20ms;
    CompletedHoldCalls : UINT := 3;
    Setup : INT := 0;
    ResetResponse : INT := 1;
    StartExecution : INT := 2;
    ReachRunning : INT := 3;
    CompleteChildren : INT := 4;
    EnterCompleting : INT := 5;
    WaitCompletion : INT := 6;
    HoldCompleted : INT := 7;
    RecoveryReset : INT := 8;
    RecoveryReady : INT := 9;
    Done : INT := 10;
END_VAR

SUPER^();

{region 'Documentation'}
(*!
<summary>Contributes only the checking Assertions, not the intentionally controlled subject results.</summary>
*)
{endregion}
METHOD PROTECTED AggregateResults
VAR_INPUT
    Aggregator : I_ResultAggregator; //! Borrowed result sink owned by the outer Test Case; add this test's checking Assertions without resetting or retaining the sink.
END_VAR
Aggregator.AddProvider(Provider := FStatePath);
Aggregator.AddProvider(Provider := FTiming);
Aggregator.AddProvider(Provider := FFinalEvents);
Aggregator.AddProvider(Provider := FPublishedPayload);
Aggregator.AddProvider(Provider := FLiveStatus);
Aggregator.AddProvider(Provider := FDiagnostics);
Aggregator.AddProvider(Provider := FChildCalls);
Aggregator.AddProvider(Provider := FRecovery);
END_METHOD

{region 'Documentation'}
(*!
<summary>Checks one final pair, immutable payloads, terminal ordering and exactly one fallback diagnostic.</summary>
*)
{endregion}
METHOD PRIVATE CheckEvents
VAR
    Index : UINT;
    ResultCount : UINT;
    AggregationCount : UINT;
    CompletedCount : UINT;
    DiagnosticCount : UINT;
    ExpectedDiagnostics : UINT;
    CompletedSequence : UDINT;
    DiagnosticSequence : UDINT;
    ExpectedMessage : STRING(GVL_Constants.MessageLength);
    ExpectedSeverity : E_EventSeverity;
END_VAR
FFinalEventsMatches := TRUE;
FPublishedPayloadMatches := TRUE;
FDiagnosticsMatches := TRUE;
FOR Index := 1 TO FCaptureFifo.ElementCount DO
    IF FEvents[Index].Name <> FSubject.Name THEN
        FFinalEventsMatches := FALSE;
        CONTINUE;
    END_IF;
    CASE FEvents[Index].EventType OF
        E_EventType.Result:
            ResultCount := ResultCount + 1;
            IF FPublishedResult.SequenceId = 0 THEN
                FPublishedResult := FEvents[Index];
            END_IF;
            FPublishedPayloadMatches := FPublishedPayloadMatches
                AND IsEventUnchanged(Event := FEvents[Index],
                    Published := FPublishedResult);
        E_EventType.Aggregation:
            AggregationCount := AggregationCount + 1;
            IF FPublishedAggregation.SequenceId = 0 THEN
                FPublishedAggregation := FEvents[Index];
            END_IF;
            FPublishedPayloadMatches := FPublishedPayloadMatches
                AND IsEventUnchanged(Event := FEvents[Index],
                    Published := FPublishedAggregation);
        E_EventType.StateTransition:
            IF FEvents[Index].State = E_State.Completed THEN
                CompletedCount := CompletedCount + 1;
                CompletedSequence := FEvents[Index].SequenceId;
            END_IF;
        E_EventType.Framework:
            DiagnosticCount := DiagnosticCount + 1;
            DiagnosticSequence := FEvents[Index].SequenceId;
            FDiagnosticsMatches := FDiagnosticsMatches
                AND (FEvents[Index].Severity = E_EventSeverity.Error);
            IF Scenario = E_RunControlCompletionScenario.InvalidTime THEN
                FDiagnosticsMatches := FDiagnosticsMatches AND (FEvents[Index].State = E_State.Completing);
            ELSIF Scenario = E_RunControlCompletionScenario.LateResetChildren THEN
                FDiagnosticsMatches := FDiagnosticsMatches AND (FEvents[Index].State = E_State.Reset);
            ELSE
                FDiagnosticsMatches := FALSE;
            END_IF;
    END_CASE;
END_FOR;
ExpectedMessage := 'Run completed.';
ExpectedSeverity := E_EventSeverity.Info;
IF FExpectedResult = E_Result.Error THEN
    ExpectedMessage := 'Run completed with error.';
    ExpectedSeverity := E_EventSeverity.Error;
END_IF;
FPublishedPayloadMatches := FPublishedPayloadMatches
    AND (FPublishedResult.Message = ExpectedMessage)
    AND (FPublishedResult.OwnerScope = E_OwnerScope.RunControl)
    AND (FPublishedResult.ResourceName = 'Fixture')
    AND (FPublishedResult.Result = FExpectedResult)
    AND (FPublishedResult.State = E_State.Completing)
    AND (FPublishedResult.Severity = ExpectedSeverity)
    AND (FPublishedAggregation.OwnerScope = E_OwnerScope.RunControl)
    AND (FPublishedAggregation.ResourceName = '')
    AND (FPublishedAggregation.Result = FExpectedResult)
    AND (FPublishedAggregation.State = E_State.Completing)
    AND (FPublishedAggregation.Severity = ExpectedSeverity);
IF Scenario = E_RunControlCompletionScenario.LateResetChildren THEN
    ExpectedMessage := '{"total":2,"inactive":0,"idle":0,"running":0,"completed":0,"passed":0,"failed":0,"error":0,"runtime":';
ELSE
    ExpectedMessage := '{"total":2,"inactive":0,"idle":0,"running":0,"completed":2,"passed":2,"failed":0,"error":0,"runtime":';
END_IF;
ExpectedMessage := CONCAT(ExpectedMessage, UDINT_TO_STRING(TIME_TO_UDINT(FFinalRuntime)));
ExpectedMessage := CONCAT(ExpectedMessage, ',"lostEvents":0}');
FPublishedPayloadMatches := FPublishedPayloadMatches AND (FPublishedAggregation.Message = ExpectedMessage);
FFinalEventsMatches := FFinalEventsMatches AND (ResultCount = 1) AND (AggregationCount = 1)
    AND (FPublishedResult.SequenceId < FPublishedAggregation.SequenceId)
    AND (CompletedCount = BOOL_TO_UINT(FSubject.IsComplete))
    AND (FCaptureStatus.LostEventCount = 0);
IF FSubject.IsComplete THEN
    FFinalEventsMatches := FFinalEventsMatches AND (FPublishedAggregation.SequenceId < CompletedSequence);
END_IF;
IF Scenario = E_RunControlCompletionScenario.LateResetChildren THEN
    ExpectedDiagnostics := 1;
ELSIF (Scenario = E_RunControlCompletionScenario.InvalidTime) AND (FStep >= WaitCompletion) THEN
    ExpectedDiagnostics := 1;
    FDiagnosticsMatches := FDiagnosticsMatches
        AND (FPublishedAggregation.SequenceId < DiagnosticSequence)
        AND (DiagnosticSequence < CompletedSequence);
END_IF;
FDiagnosticsMatches := FDiagnosticsMatches AND (DiagnosticCount = ExpectedDiagnostics);
END_METHOD

{region 'Documentation'}
(*!
<summary>Initializes the checking Assertions; the scenario explicitly initializes its isolated subject.</summary>
*)
{endregion}
METHOD PROTECTED Configure
FPreparationStateCount := 0;
FTestStateCount := 1;
FStatePath.Initialize(Parent := THIS^,
    AssertionName := 'StatePath');
FTiming.Initialize(Parent := THIS^,
    AssertionName := 'Timing');
FFinalEvents.Initialize(Parent := THIS^,
    AssertionName := 'FinalEvents');
FPublishedPayload.Initialize(Parent := THIS^,
    AssertionName := 'PublishedPayload');
FLiveStatus.Initialize(Parent := THIS^,
    AssertionName := 'LiveStatus');
FDiagnostics.Initialize(Parent := THIS^,
    AssertionName := 'Diagnostics');
FChildCalls.Initialize(Parent := THIS^,
    AssertionName := 'ChildCalls');
FRecovery.Initialize(Parent := THIS^,
    AssertionName := 'Recovery');
END_METHOD

{region 'Documentation'}
(*!
<summary>Compares captured event fields explicitly, without relying on structure padding.</summary>
*)
{endregion}
METHOD PRIVATE IsEventUnchanged : BOOL //! TRUE when all defined event fields match the retained snapshot; structure padding is ignored.
VAR_IN_OUT CONSTANT
    Event : ST_Event; //! Borrowed read-only event to compare field by field.
    Published : ST_Event; //! Borrowed read-only publication snapshot used as the expected value.
END_VAR
IsEventUnchanged := (Event.SequenceId = Published.SequenceId)
    AND (Event.Timestamp = Published.Timestamp)
    AND (Event.OwnerScope = Published.OwnerScope)
    AND (Event.EventType = Published.EventType)
    AND (Event.Severity = Published.Severity)
    AND (Event.Name = Published.Name)
    AND (Event.ResourceName = Published.ResourceName)
    AND (Event.State = Published.State)
    AND (Event.Result = Published.Result)
    AND (Event.Message = Published.Message);
END_METHOD

{region 'Documentation'}
(*!
<summary>No asynchronous test resource remains to stop.</summary>
*)
{endregion}
METHOD PROTECTED ProcessAbort
VAR_INPUT
    Enable : BOOL; //! Phase permission supplied by the owning Test Case; FALSE does not authorize progression, while observation may continue.
END_VAR
IF Enable THEN
    CompleteAbort();
END_IF;
END_METHOD

{region 'Documentation'}
(*!
<summary>Checks each subject call before allowing the script to advance; failures remain latched.</summary>
*)
{endregion}
METHOD PROTECTED ProcessAssertions
VAR_INPUT
    Enable : BOOL; //! Phase permission supplied by the owning Test Case; FALSE does not authorize progression, while observation may continue.
END_VAR
FStatePath(Enable := Enable,
    State := State,
    IN := FStatePathMatches);
FTiming(Enable := Enable,
    State := State,
    IN := FTimingMatches);
FFinalEvents(Enable := Enable,
    State := State,
    IN := FFinalEventsMatches);
FPublishedPayload(Enable := Enable,
    State := State,
    IN := FPublishedPayloadMatches);
FLiveStatus(Enable := Enable,
    State := State,
    IN := FLiveStatusMatches);
FDiagnostics(Enable := Enable,
    State := State,
    IN := FDiagnosticsMatches);
FChildCalls(Enable := Enable,
    State := State,
    IN := FChildCallsMatches);
FRecovery(Enable := Enable,
    State := State,
    IN := FRecoveryMatches);
IF Enable THEN
    FStepChecked := TRUE;
END_IF;
END_METHOD

{region 'Documentation'}
(*!
<summary>No resource Preparation is required for this controlled owner scenario.</summary>
*)
{endregion}
METHOD PROTECTED ProcessPreparations
VAR_INPUT
    // SA0033: Required override; the scenario has no Preparation phase.
    {attribute 'analysis' := '-33'}
    Enable : BOOL; //! Phase permission supplied by the owning Test Case; FALSE does not authorize progression, while observation may continue.
END_VAR
END_METHOD

{region 'Documentation'}
(*!
<summary>Restarts the test script and clears checking Assertions; subject setup belongs to the next test attempt.</summary>
*)
{endregion}
METHOD PROTECTED ProcessReset
FStep := Setup;
FNextStep := Setup;
FStepChecked := FALSE;
FCallCount := 0;
FEntryCall := 0;
FHoldCalls := 0;
FPublishedResult.SequenceId := 0;
FPublishedAggregation.SequenceId := 0;
FDelayClock.Reset();
FStatePathMatches := TRUE;
FTimingMatches := TRUE;
FFinalEventsMatches := TRUE;
FPublishedPayloadMatches := TRUE;
FLiveStatusMatches := TRUE;
FDiagnosticsMatches := TRUE;
FChildCallsMatches := TRUE;
FRecoveryMatches := TRUE;
FStatePath.Reset();
FTiming.Reset();
FFinalEvents.Reset();
FPublishedPayload.Reset();
FLiveStatus.Reset();
FDiagnostics.Reset();
FChildCalls.Reset();
FRecovery.Reset();
CompleteReset();
END_METHOD

{region 'Documentation'}
(*!
<summary>Advances the explicit test script with at most one subject FB call per active PLC cycle.</summary>
*)
{endregion}
METHOD PROTECTED ProcessTests
VAR_INPUT
    Enable : BOOL; //! Phase permission supplied by the owning Test Case; FALSE does not authorize progression, while observation may continue.
END_VAR
IF NOT Enable THEN
    RETURN;
END_IF;
IF FStepChecked THEN
    FStep := FNextStep;
    FStepChecked := FALSE;
END_IF;
IF FStep = Done THEN
    CompleteTests();
    RETURN;
END_IF;
RunStep();
END_METHOD

{region 'Documentation'}
(*!
<summary>Arranges one call and compares timing, state, publication and cyclic observations.</summary>
*)
{endregion}
METHOD PRIVATE RunStep
VAR
    Config : ST_RunConfig;
    Snapshot : ST_RunControlStatus;
    ExpectedState : E_State;
    ExpectedResult : E_Result;
    ExpectedTask : E_OrchestratorTask;
    ExpectedCompleted : UINT;
    ExpectedPassed : UINT;
END_VAR
FDelayClock.Update();
FNextStep := FStep + 1;
ExpectedResult := E_Result.NotEvaluated;
ExpectedTask := E_OrchestratorTask.Idle;

CASE FStep OF
    Setup:
        FDelay := DefaultDelay;
        FExpectedResult := E_Result.Passed;
        FTimingMatches := Config.CompletionDelay = DefaultDelay;
        IF Scenario = E_RunControlCompletionScenario.ZeroDelay THEN
            Config.CompletionDelay := T#0ms;
            FDelay := T#0ms;
        END_IF;
        IF Scenario = E_RunControlCompletionScenario.LateResetChildren THEN
            Config.ResetTimeout := ResetDeadline;
            FExpectedResult := E_Result.Error;
        END_IF;
        IF NOT FCapture.Initialize(Buffer := FEvents,
            FifoControl := FCaptureFifo,
            Status := FCaptureStatus) THEN
            Error(Message := 'Completion capture could not be initialized.');
            RETURN;
        END_IF;
        FHelper.BeginScenario();
        FSubject.Bind(Publisher := FCapture,
            Helper := FHelper,
            Config := Config);
        IF NOT FSubject.Initialize(Name := 'CompletionSubject',
            EventBuffer := FCapture) THEN
            Error(Message := 'Completion subject could not be initialized.');
            RETURN;
        END_IF;
        FFirstChild.State := E_State.Reset;
        FFirstChild.Ready := FALSE;
        FFirstChild.Complete := FALSE;
        FFirstChild.Result := E_Result.NotEvaluated;
        FSecondChild := FFirstChild;
        ExpectedState := E_State.Reset;
        ExpectedTask := E_OrchestratorTask.Reset;

    ResetResponse:
        IF Scenario = E_RunControlCompletionScenario.LateResetChildren THEN
            // The root deadline expires while children are still resetting.
            ExpectedState := E_State.Reset;
            ExpectedTask := E_OrchestratorTask.Reset;
            FNextStep := ResetResponse;
        ELSE
            FHelper.SetObservation(Ready := TRUE,
                ResetFinished := TRUE);
            FFirstChild.State := E_State.Idle;
            FFirstChild.Ready := TRUE;
            FSecondChild := FFirstChild;
            ExpectedState := E_State.Idle;
        END_IF;

    StartExecution:
        FSubject.RequestStart();
        FFirstChild.State := E_State.Running;
        FFirstChild.Ready := FALSE;
        FSecondChild := FFirstChild;
        ExpectedState := E_State.Starting;
        ExpectedTask := E_OrchestratorTask.Execution;

    ReachRunning:
        FHelper.SetObservation(Ready := FALSE);
        ExpectedState := E_State.Running;
        ExpectedTask := E_OrchestratorTask.Execution;

    CompleteChildren:
        FFirstChild.State := E_State.Completed;
        FFirstChild.Result := E_Result.Passed;
        FFirstChild.Complete := TRUE;
        FSecondChild := FFirstChild;
        ExpectedState := E_State.Running;
        ExpectedTask := E_OrchestratorTask.Execution;

    EnterCompleting:
        FHelper.SetObservation(Ready := FALSE,
            ExecutionFinished := TRUE);
        ExpectedState := E_State.Completing;
        ExpectedResult := FExpectedResult;
        ExpectedTask := E_OrchestratorTask.Execution;

    WaitCompletion:
        IF Scenario = E_RunControlCompletionScenario.InvalidTime THEN
            FSubject.SetInvalidCompletionTime(Invalid := TRUE);
        END_IF;
        IF Scenario = E_RunControlCompletionScenario.LateResetChildren THEN
            FFirstChild.State := E_State.Completed;
            FFirstChild.Result := E_Result.Error;
            FFirstChild.Complete := TRUE;
            // Only this child finishes during the delay; the second finishes after Completed.
        END_IF;
        ExpectedState := E_State.Completing;
        ExpectedResult := FExpectedResult;
        ExpectedTask := E_OrchestratorTask.Execution;
        IF Scenario = E_RunControlCompletionScenario.LateResetChildren THEN
            ExpectedTask := E_OrchestratorTask.Idle;
        END_IF;
        IF (Scenario = E_RunControlCompletionScenario.InvalidTime)
            OR (FDelayClock.ElapsedLTime >= TIME_TO_LTIME(FDelay)) THEN
            ExpectedState := E_State.Completed;
            ExpectedTask := E_OrchestratorTask.Idle;
        ELSE
            FNextStep := WaitCompletion;
        END_IF;

    HoldCompleted:
        IF Scenario = E_RunControlCompletionScenario.LateResetChildren THEN
            FSecondChild.State := E_State.Completed;
            FSecondChild.Result := E_Result.Passed;
            FSecondChild.Complete := TRUE;
        END_IF;
        ExpectedState := E_State.Completed;
        ExpectedResult := FExpectedResult;
        FHoldCalls := FHoldCalls + 1;
        IF FHoldCalls < CompletedHoldCalls THEN
            FNextStep := HoldCompleted;
        END_IF;

    RecoveryReset:
        FSubject.SetInvalidCompletionTime(Invalid := FALSE);
        FHelper.SetObservation(Ready := FALSE);
        FSubject.RequestReset();
        FFirstChild.State := E_State.Reset;
        FFirstChild.Result := E_Result.NotEvaluated;
        FFirstChild.Complete := FALSE;
        FFirstChild.Ready := FALSE;
        FSecondChild := FFirstChild;
        ExpectedState := E_State.Reset;
        ExpectedTask := E_OrchestratorTask.Reset;

    RecoveryReady:
        FHelper.SetObservation(Ready := TRUE,
            ResetFinished := TRUE);
        FFirstChild.State := E_State.Idle;
        FFirstChild.Ready := TRUE;
        FSecondChild := FFirstChild;
        ExpectedState := E_State.Idle;
ELSE
    Error(Message := 'Unexpected completion test step.');
    RETURN;
END_CASE;

FSubject.SetChildObservations(FirstChild := FFirstChild,
    SecondChild := FSecondChild);
FSubject(ControlData := FControl);
FCallCount := FCallCount + 1;
Snapshot := FSubject.Status;

IF (FStep = ResetResponse) AND (Scenario = E_RunControlCompletionScenario.LateResetChildren)
    AND (FSubject.State = E_State.Completing) THEN
    ExpectedState := E_State.Completing;
    ExpectedResult := E_Result.Error;
    ExpectedTask := E_OrchestratorTask.Idle;
    FNextStep := WaitCompletion;
END_IF;
IF (ExpectedState = E_State.Completing) AND (FEntryCall = 0) THEN
    FEntryCall := FCallCount;
    FDelayClock.Start();
    FFinalRuntime := Snapshot.Runtime;
END_IF;

FStatePathMatches := (FSubject.State = ExpectedState)
    AND (Snapshot.Execution.State = ExpectedState)
    AND (FControl.Status.Execution.State = ExpectedState)
    AND (FSubject.Result = ExpectedResult)
    AND (FControl.Status.Execution.Result = ExpectedResult)
    AND (FHelper.CurrentTask = ExpectedTask);
FChildCallsMatches := (FSubject.ChildCallCount = FCallCount)
    AND FSubject.ChildBodyCallsMatch
    AND (FHelper.ExecuteCount = FCallCount);

IF (FStep = WaitCompletion) OR (FStep = HoldCompleted) THEN
    FTimingMatches := FDelayClock.IsValid AND (FCallCount > FEntryCall)
        AND (Snapshot.Runtime = FFinalRuntime);
    IF Scenario <> E_RunControlCompletionScenario.InvalidTime THEN
        FTimingMatches := FTimingMatches
            AND ((FSubject.State = E_State.Completed)
                = (FDelayClock.ElapsedLTime >= TIME_TO_LTIME(FDelay)));
    END_IF;
    FLiveStatusMatches := Snapshot.SuiteCountTotal = 2;
    IF Scenario = E_RunControlCompletionScenario.LateResetChildren THEN
        ExpectedCompleted := 1;
        ExpectedPassed := 0;
        IF FStep = HoldCompleted THEN
            ExpectedCompleted := 2;
            ExpectedPassed := 1;
        END_IF;
        FLiveStatusMatches := FLiveStatusMatches
            AND (Snapshot.SuiteCountCompleted = ExpectedCompleted)
            AND (Snapshot.SuiteCountPassed = ExpectedPassed)
            AND (Snapshot.SuiteCountError = 1)
            AND (FControl.Status.SuiteCountCompleted = ExpectedCompleted)
            AND (FControl.Status.SuiteCountPassed = ExpectedPassed);
    ELSE
        FLiveStatusMatches := FLiveStatusMatches
            AND (Snapshot.SuiteCountCompleted = 2) AND (Snapshot.SuiteCountPassed = 2);
    END_IF;
END_IF;
IF (FEntryCall > 0) AND (FStep < RecoveryReset) THEN
    CheckEvents();
END_IF;
IF FStep = RecoveryReady THEN
    FRecoveryMatches := FSubject.IsReady AND (FSubject.Result = E_Result.NotEvaluated)
        AND NOT FSubject.HasResetTimeout AND NOT FSubject.HasTimeout AND NOT FSubject.HasAbortTimeout
        AND (FSubject.ConfigureCount = 1) AND (FHelper.InitializeCount = 1);
END_IF;
END_METHOD

END_FUNCTION_BLOCK

// ---- SelfTests/TestSuites/TestSuite_CommandAdapter.TcPOU
{region 'Documentation'}
(*!
<summary>Groups isolated command-adapter initialization, qualification and field-independence tests.</summary>
*)
{endregion}
FUNCTION_BLOCK TestSuite_CommandAdapter EXTENDS TestSuiteBase
VAR
    FInitialization : Test_CommandAdapterInitialization;
    FReinitialization : Test_CommandAdapterInitialization;
    FStartQualification : Test_CommandQualification;
    FAbortQualification : Test_CommandQualification;
    FResetQualification : Test_CommandQualification;
    FIndependentCommands : Test_CommandIndependence;
    FTestCases : ARRAY[1..TestCaseCapacity] OF I_TestCase;
END_VAR
VAR CONSTANT
    TestCaseCapacity : UINT := 6;
END_VAR

SUPER^();

{region 'Documentation'}
(*!
<summary>Initializes and registers the local command scenarios for serial execution.</summary>
*)
{endregion}
METHOD PROTECTED Configure
VAR_IN_OUT
    // SA0167: Borrowed owner builder; no temporary instance is created.
    {attribute 'analysis' := '-167'}
    Builder : TestSuiteConfigurationBuilder; //! Borrowed owner configuration builder used only during this Configure call; register this owner's concrete children.
END_VAR
VAR
    TestConfig : ST_TestCaseConfig;
END_VAR
Builder.Initialize(Mode := E_OrchestrationMode.Serial,
    TestCases := FTestCases);
FInitialization.Initialize(Parent := THIS^,
    TestName := 'Initialization',
    Config := TestConfig);
Builder.Register(TestCase := FInitialization);
FReinitialization.Initialize(Parent := THIS^,
    TestName := 'Reinitialization',
    Config := TestConfig);
Builder.Register(TestCase := FReinitialization);
FStartQualification.Initialize(Parent := THIS^,
    TestName := 'StartQualification',
    Config := TestConfig);
Builder.Register(TestCase := FStartQualification);
FAbortQualification.Initialize(Parent := THIS^,
    TestName := 'AbortQualification',
    Config := TestConfig);
Builder.Register(TestCase := FAbortQualification);
FResetQualification.Initialize(Parent := THIS^,
    TestName := 'ResetQualification',
    Config := TestConfig);
Builder.Register(TestCase := FResetQualification);
FIndependentCommands.Initialize(Parent := THIS^,
    TestName := 'IndependentCommands',
    Config := TestConfig);
Builder.Register(TestCase := FIndependentCommands);
END_METHOD

{region 'Documentation'}
(*!
<summary>Returns a registered scenario using its original array index.</summary>
*)
{endregion}
METHOD PUBLIC GetTestCase : I_TestCase //! Typed child interface at the original array index; zero when no entry is available.
VAR_INPUT
    Index : DINT; //! Original occupied child-array index, rather than an ordinal position.
END_VAR
GetTestCase := 0;
IF (ChildCount = 0) OR (Index < ChildArrayLowerBound)
    OR (DINT_TO_LINT(Index) >= DINT_TO_LINT(ChildArrayLowerBound) + UINT_TO_LINT(ChildCount)) THEN
    RETURN;
END_IF;
GetTestCase := FTestCases[Index];
END_METHOD

{region 'Documentation'}
(*!
<summary>Calls each owned scenario once per initialized Suite cycle.</summary>
*)
{endregion}
METHOD PROTECTED ProcessTestCases
FInitialization(PrimeHistory := FALSE);
FReinitialization(PrimeHistory := TRUE);
FStartQualification(Command := E_AdapterCommand.Start);
FAbortQualification(Command := E_AdapterCommand.Abort);
FResetQualification(Command := E_AdapterCommand.Reset);
FIndependentCommands();
END_METHOD

END_FUNCTION_BLOCK

